(* IEC 61131-3 sources: daoli-st-library/DL_Algo (part 20) *)

(* ---- FB_DL_ResonanceTrackNotch.st ---- *)
(*
  FB_DL_ResonanceTrackNotch  —  共振频率跟踪与陷波中心估计 / Resonance frequency tracking and notch centre estimation
  分类 Category : DL_Algo
  码位 Code     : 16#02_3_82
  版本 Version  : 1.0.1
  来源 Source   : t1-6-plcopen — IEC 61131-3 标准语义的道莅防御性实现
  溯源 Origin   : PLCopen 运动/振动监视公开语义借鉴，clean-room 实现，仅借分类与参数域，未复制任何源码行
  功能 Function : 1) 二阶带通相位过零测周期：以信号上行过零点之间的累计时间为一个周期 [s]，取倒数得频率 [Hz]；
                  2) 频率估计经 5 点滑动中值去野值（排序网络，无循环），抗单点脉冲干扰；
                  3) 中值结果钳制到 [fFreqMinHz, fFreqMaxHz]，输出 fResonanceHz 供陷波中心使用；
                  4) 连续 nSettleCycles 次估计落在中心 ±fLockBandHz 内 → bLocked；锁定后须连续
                     nLostCycles 次越带才降级（迟滞，防抖）；
                  5) fTrackConfidence 逐拍升降（步长 DL_CONF_STEP），幅值不足时衰减而非清零。
  边界 Boundary : ① fSampleDt <= 0 / 搜索窗倒置 / 搜索窗越奈奎斯特（fFreqMaxHz >= 1/(2·fSampleDt)）
                     任一成立判组态错置 0382，状态进 eFault 且不投运（R28 组态域闸覆盖全部换算引脚）；
                  ② 信号幅值（峰值包络）< fAmpFloor 时不出频率结论：bLocked := FALSE，估计值保持，
                     置信度按 DL_CONF_DECAY 衰减（不置 bError，信息级 01B2，R187③）；
                  ③ 频率跳变率超 fMaxSlewHzPerSec 判野值丢弃并计数；计数在 DL_WILD_WINDOW 窗内
                     超 nWildMax 置「跟踪发散」故障 0392（计数窗由自复位 TON 滚动清零）；
                  ④ 幅值门限只影响结论不影响估计：无结论期间 fResonanceHz 保持末次有效值（R191 显式声明）；
                  ⑤ 解除路径自证：_bFault 清除 = rtReset.Q 单一路径（引脚可满足）；发散码 0392 另可由
                     「窗内野值计数回落至 0」按码专清（两路径互不掩盖）。
  依赖 Depends  : 仅 Standard.library（TON / R_TRIG / ABS / MAX / MIN / MOD），零外部组件依赖
  同拍双窗配比  : 野值观察窗 DL_WILD_WINDOW = 2 s 与锁定计数 nSettleCycles ≥ 1 不同源；
                  配比约束 nSettleCycles × fSampleDt <= DL_WILD_WINDOW，保证锁定判据至少跨一个观察窗成立

  码表 Error codes（本件格 02_3_82，子码步进 +0x10）:
    16#0002_0382 故障级：组态非法（采样周期 <= 0 / 搜索窗倒置 / 越奈奎斯特 / 锁定带或幅值下限 <= 0）
    16#0002_0392 故障级：跟踪发散（野值计数超 nWildMax，跟踪环已失去物理意义）
    16#0002_03A2 故障级：状态机落 ELSE 兜底（非法相位 ID）
    16#0002_01B2 信息级：信号幅值低于 fAmpFloor，本拍不出频率结论（不置 bError）
    16#0002_01C2 信息级：单拍野值已丢弃（跳变率超 fMaxSlewHzPerSec，不置 bError）

  修订历史 Revision :
    2026-11-18  v1.0.0  R37 首版
  修订 History : v1.0.1 2026-11-18 R37 终审：锁定出口随幅值门限/保持相同拍降级（原缺 eTrack/eHold 分支归零）
*)

TYPE E_DL_ResTrackState :
(
    eIdle     := 0,   // 空闲：未使能，不出结论 / Idle, no conclusion while disabled
    eTrack    := 10,  // 跟踪中：已取得周期，尚未满足锁定次数 / Tracking, period acquired but lock count insufficient
    eLocked   := 20,  // 已锁定：连续在带次数达标 / Locked, the in-band count reached the preset
    eHold     := 30,  // 保持：幅值不足，估计保持、置信度衰减 / Hold, low amplitude, estimate held and confidence decaying
    eDiverged := 40,  // 发散：野值计数超限，跟踪失效 / Diverged, wild-value count exceeded
    eFault    := 90   // 故障：组态非法或状态兜底锁定 / Fault, illegal configuration or fallback
);
END_TYPE

FUNCTION_BLOCK FB_DL_ResonanceTrackNotch
VAR_INPUT
    bEnable        : BOOL := FALSE;              // 总使能，FALSE 时不出结论并回 eIdle / Master enable
    bReset         : BOOL := FALSE;              // 复位，上升沿清故障锁存 / Reset, rising edge clears the fault latch
    fSignal        : REAL := 0.0;                // 振动或电流反馈原始信号 [工程单位] / Raw vibration or current feedback
    fSampleDt      : REAL := 0.010;              // 采样周期 [s]，域 > 0 / Sampling period [s], domain > 0
    fFreqMinHz     : REAL := 20.0;               // 搜索窗下限 [Hz]，域 > 0 / Search window lower limit [Hz]
    fFreqMaxHz     : REAL := 400.0;              // 搜索窗上限 [Hz]，须 > 下限且 < 奈奎斯特 / Search window upper limit [Hz]
    fLockBandHz    : REAL := 2.0;                // 锁定带宽（中心 ± 本值）[Hz]，域 > 0 / Lock band half width [Hz]
    fAmpFloor      : REAL := 0.05;               // 幅值下限，低于此不出结论 [工程单位]，域 > 0 / Amplitude floor
    fMaxSlewHzPerSec : REAL := 500.0;            // 允许最大频率跳变率 [Hz/s]，域 > 0 / Permitted frequency slew [Hz/s]
    nSettleCycles  : INT := 5;                   // 连续在带次数门限 [次]，域 >= 1 / In-band settle cycles
    nLostCycles    : INT := 3;                   // 连续越带次数门限（迟滞）[次]，域 >= 1 / Out-of-band lost cycles
    nWildMax       : INT := 8;                   // 窗内野值计数上限 [次]，超过即判发散 / Wild-value count limit
END_VAR
VAR_OUTPUT
    fResonanceHz     : REAL;                     // 共振频率估计（钳制后、去野值）[Hz] / Resonance frequency estimate [Hz]
    fTrackConfidence : REAL;                     // 跟踪置信度 [0~1 无量纲] / Tracking confidence, 0..1
    bLocked          : BOOL;                     // 锁定标志（迟滞维持）/ Locked flag with hysteresis
    bValid           : BOOL;                     // 本拍估计可用标志 / Estimate usable this scan
    bError           : BOOL;                     // 故障标志，派生自锁存 / Fault flag derived from the latch
    nErrId           : UDINT;                    // 事件码，0 = 无事件 / Event code, 0 = no event
    eStateOut        : E_DL_ResTrackState;       // 状态出口，段尾单点映射 / State outlet, mapped at the tail
END_VAR
VAR
    tonWild        : TON;                        // 野值观察窗，自复位（IN := NOT Q）/ Wild-value observation window, self-resetting
    rtReset        : R_TRIG;                     // 复位上升沿 / Reset rising edge
    rtEnable       : R_TRIG;                     // 使能上升沿 / Enable rising edge
    _eState        : E_DL_ResTrackState := E_DL_ResTrackState.eIdle;  // 内部相位（CASE 只写本量）/ Internal phase, the only CASE target
    _uFault        : UDINT;                      // 故障码锁存（仅复位沿或按码专清）/ Latched fault code
    _uInfo         : UDINT;                      // 信息码，每拍重算 / Information code, recomputed per scan
    _bFault        : BOOL;                       // 故障锁存位 / Latched fault bit
    _bCfgBad       : BOOL;                       // 组态非法聚合 / Configuration invalid aggregate
    _bAmpLow       : BOOL;                       // 幅值不足判定 / Low amplitude predicate
    _bWildScan     : BOOL;                       // 本拍野值丢弃标志 / Wild value discarded this scan
    _bCrossUp      : BOOL;                       // 上行过零事件 / Upward zero-crossing event
    _bHavePeriod   : BOOL;                       // 已捕获至少一个完整周期 / At least one full period captured
    fSignalPrev    : REAL;                       // 上拍信号快照 [工程单位] / Previous-scan signal snapshot
    fCrossAccum    : REAL;                       // 过零后累计时间 [s] / Elapsed time since the last up-crossing [s]
    fPeriodSec     : REAL;                       // 实测周期 [s] / Measured period [s]
    fFreqRaw       : REAL;                       // 单次频率估计（未去野）[Hz] / Raw frequency estimate [Hz]
    fFreqMed       : REAL;                       // 中值去野后的频率 [Hz] / Median-filtered frequency [Hz]
    fFreqAcc       : REAL;                       // 已受理的频率（钳制后）[Hz] / Accepted frequency after clamping [Hz]
    fFreqPrev      : REAL;                       // 上一个已受理频率（跳变率基准）[Hz] / Previous accepted frequency [Hz]
    fCenterHz      : REAL;                       // 锁定中心频率 [Hz] / Lock centre frequency [Hz]
    fAmpEnv        : REAL;                       // 峰值包络（带衰减）[工程单位] / Decaying peak envelope
    fConfidence    : REAL := 0.0;                // 置信度保持量 [0~1] / Held confidence value
    afFreqBuf      : ARRAY[0..4] OF REAL;        // 5 点滑动缓冲 [Hz] / Five-point sliding buffer [Hz]
    nBufIdx        : INT;                        // 缓冲写指针 [索引] / Buffer write index
    nFill          : INT;                        // 缓冲已填点数 [个] / Filled slots in the buffer
    nInBandCnt     : INT;                        // 连续在带计数 [次] / Consecutive in-band count
    nOutBandCnt    : INT;                        // 连续越带计数 [次] / Consecutive out-of-band count
    nWildCnt       : INT;                        // 窗内野值计数 [次] / Wild-value count inside the window
    fSort0         : REAL;                       // 排序中间量 0 [Hz] / Sorting scratch 0 [Hz]
    fSort1         : REAL;                       // 排序中间量 1 [Hz] / Sorting scratch 1 [Hz]
    fSort2         : REAL;                       // 排序中间量 2 [Hz] / Sorting scratch 2 [Hz]
    fSort3         : REAL;                       // 排序中间量 3 [Hz] / Sorting scratch 3 [Hz]
    fSort4         : REAL;                       // 排序中间量 4 [Hz] / Sorting scratch 4 [Hz]
    fSwap          : REAL;                       // 排序交换临时量 [Hz] / Sorting swap scratch [Hz]
END_VAR
VAR CONSTANT
    DL_WILD_WINDOW : TIME  := T#2S;      // 野值观察窗 [ms]，自复位节拍 / Wild-value window, self-resetting
    DL_WILD_WINDOW_SEC : REAL := 2.0;    // 野值观察窗秒值 [s]，与上行同源 / Wild-value window in seconds
    DL_NYQ_RATIO   : REAL  := 0.5;       // 奈奎斯特系数（fs/2）[1] / Nyquist factor
    DL_CONF_STEP   : REAL  := 0.05;      // 置信度上升步长 [1/拍] / Confidence rising step
    DL_CONF_DECAY  : REAL  := 0.90;      // 低幅值衰减系数 [1/拍] / Confidence decay factor under low amplitude
    DL_AMP_DECAY   : REAL  := 0.95;      // 峰值包络衰减系数 [1/拍] / Peak envelope decay factor
    DL_EPS         : REAL  := 1.0E-6;    // 判零容差 [1] / Zero tolerance
    DL_BUF_LEN     : INT   := 5;         // 滑动缓冲长度 [个] / Sliding buffer length
END_VAR

(* —— 段 0：边缘检测与自复位节拍窗无条件周期刷新（禁置于任何分支内，R182） —— *)
rtReset(CLK := bReset);                                          // 复位上升沿，每拍必调 / Reset edge, called every scan
rtEnable(CLK := bEnable);                                        // 使能上升沿，每拍必调 / Enable edge, called every scan
tonWild(IN := NOT tonWild.Q, PT := DL_WILD_WINDOW);              // 野值窗自复位：到点后下一拍断输入归零 / Self-resetting window

(* —— 段 1：单拍量预清零（快照 / 锁存 / 计数不入清单，R187①） —— *)
_uInfo         := 16#0000_0000;   // 信息码每拍重算 / Info code recomputed
bError         := FALSE;          // 故障出口每拍重算，段 6 由锁存派生 / Fault outlet recomputed, derived in segment 6
bValid         := FALSE;          // 可用标志缺省 FALSE / Usable flag defaults FALSE
bLocked        := FALSE;          // 锁定出口缺省 FALSE / Locked outlet defaults FALSE
_bCfgBad       := FALSE;          // 组态非法聚合预清零 / Config aggregate pre-cleared
_bAmpLow       := FALSE;          // 低幅值判定预清零 / Low amplitude pre-cleared
_bWildScan     := FALSE;          // 本拍野值标志预清零 / Wild flag pre-cleared
_bCrossUp      := FALSE;          // 过零事件预清零 / Crossing event pre-cleared

(* —— 段 2：复位沿清锁存 + 按码专清（R188 双路径，互不掩盖） —— *)
IF rtReset.Q THEN
    _bFault  := FALSE;            // 复位沿清锁存位 / Clear the latched bit
    _uFault  := 16#0000_0000;     // 复位沿清锁存码 / Clear the latched code
    nWildCnt := 0;                // 复位沿同步清野值计数（发散判据的输入）/ Wild count cleared with the reset
    nInBandCnt := 0;              // 复位沿清在带计数，重新建立锁 / In-band count cleared
    nOutBandCnt := 0;             // 复位沿清越带计数 / Out-of-band count cleared
    fConfidence := 0.0;           // 复位沿置信度清零 / Confidence cleared
END_IF
IF tonWild.Q THEN
    IF nWildCnt > 0 THEN
        nWildCnt := nWildCnt - 1; // 窗到点衰减一个野值（迟滞释放，避免长期积压）/ Decay one wild value per window
    END_IF
END_IF
IF (_uFault = 16#0002_0392) AND (nWildCnt = 0) THEN
    _uFault := 16#0000_0000;      // 按码专清：发散码仅在野值窗回零时清除 / Code-specific clear for the divergence code
    _bFault := FALSE;             // 锁存位同步清 / Latched bit cleared together
END_IF

(* —— 段 3：组态域闸（覆盖全部参与换算的引脚，缺一个即该判据静默失效，R151） —— *)
IF (fSampleDt <> fSampleDt) OR (fSampleDt <= 0.0) THEN
    _bCfgBad := TRUE;             // 采样周期非法（过零计时与奈奎斯特的分母）/ Sampling period illegal
END_IF
IF (fFreqMinHz <> fFreqMinHz) OR (fFreqMinHz <= 0.0) THEN
    _bCfgBad := TRUE;             // 搜索窗下限非法 / Lower search limit illegal
END_IF
IF (fFreqMaxHz <> fFreqMaxHz) OR (fFreqMaxHz <= fFreqMinHz) THEN
    _bCfgBad := TRUE;             // 搜索窗倒置（上限须严格大于下限）/ Inverted search window
END_IF
IF (fLockBandHz <> fLockBandHz) OR (fLockBandHz <= 0.0) THEN
    _bCfgBad := TRUE;             // 锁定带宽非法（迟滞判据的分母）/ Lock band illegal
END_IF
IF (fAmpFloor <> fAmpFloor) OR (fAmpFloor <= 0.0) THEN
    _bCfgBad := TRUE;             // 幅值下限非法 / Amplitude floor illegal
END_IF
IF (fMaxSlewHzPerSec <> fMaxSlewHzPerSec) OR (fMaxSlewHzPerSec <= 0.0) THEN
    _bCfgBad := TRUE;             // 跳变率上限非法（野值判据的分母）/ Slew limit illegal
END_IF
IF nSettleCycles < 1 THEN
    _bCfgBad := TRUE;             // 锁定次数门限非法 / Settle cycles illegal
END_IF
IF nLostCycles < 1 THEN
    _bCfgBad := TRUE;             // 失锁次数门限非法 / Lost cycles illegal
END_IF
IF nWildMax < 1 THEN
    _bCfgBad := TRUE;             // 野值门限非法 / Wild limit illegal
END_IF
IF (NOT _bCfgBad) AND (fFreqMaxHz >= (DL_NYQ_RATIO / fSampleDt)) THEN
    _bCfgBad := TRUE;             // 搜索窗越奈奎斯特：fMax >= fs/2 时测周期无意义 / Window crosses Nyquist
END_IF
IF _bCfgBad THEN
    _uFault := 16#0002_0382;      // 故障级：组态非法
    _bFault := TRUE;              // 锁存位置位（复位沿可清）
    bError  := TRUE;              // 故障标志置位（R45 配对）
    _eState := E_DL_ResTrackState.eFault;  // 状态机进故障相
END_IF

(* —— 段 4：跟踪内核（仅无故障且使能时执行） —— *)
IF (NOT _bFault) AND bEnable AND (NOT _bCfgBad) THEN
    (* 4.1 峰值包络：MAX 跟随上升沿，逐拍衰减，用于幅值门限 *)
    fAmpEnv := MAX(ABS(fSignal), fAmpEnv * DL_AMP_DECAY);        // 峰值包络 [工程单位]
    _bAmpLow := (fAmpEnv < fAmpFloor);                           // 幅值不足判定

    (* 4.2 上行过零测周期：上一次过零起的累计时间即周期 *)
    _bCrossUp := (fSignalPrev < 0.0) AND (fSignal >= 0.0);       // 上行过零（含恰好落 0 的边界）
    fCrossAccum := fCrossAccum + fSampleDt;                      // 过零计时累加 [s]
    IF _bCrossUp THEN
        IF _bHavePeriod THEN
            fPeriodSec := fCrossAccum;                           // 两次上行过零之间为一个周期 [s]
            IF fPeriodSec > DL_EPS THEN
                fFreqRaw := 1.0 / fPeriodSec;                    // 倒数为频率 [Hz]（分母已判 > 容差）
                afFreqBuf[nBufIdx] := fFreqRaw;                  // 入滑动缓冲
                nBufIdx := (nBufIdx + 1) MOD DL_BUF_LEN;         // 环形指针推进（移位量已归一，禁越位宽）
                IF nFill < DL_BUF_LEN THEN
                    nFill := nFill + 1;                          // 已填点数饱和到缓冲长度
                END_IF
            END_IF
        END_IF
        fCrossAccum := 0.0;                                      // 过零后计时归零（本拍唯一清零点）
        _bHavePeriod := TRUE;                                     // 已具备周期测量能力
    END_IF
    IF fCrossAccum > (DL_WILD_WINDOW_SEC) THEN
        fCrossAccum := 0.0;                                      // 超时无过零：计时器防溢出回零（信号消失路径）
        _bHavePeriod := FALSE;                                   // 周期能力失效，等待重新建立
    END_IF
    fSignalPrev := fSignal;                                      // 信号快照更新（末行，不预清零）

    (* 4.3 5 点滑动中值：排序网络（9 次比较交换），无循环 *)
    IF nFill >= DL_BUF_LEN THEN                                  // 满窗才出中值
        fSort0 := afFreqBuf[0];                                  // 拷贝 0
        fSort1 := afFreqBuf[1];                                  // 拷贝 1
        fSort2 := afFreqBuf[2];                                  // 拷贝 2
        fSort3 := afFreqBuf[3];                                  // 拷贝 3
        fSort4 := afFreqBuf[4];                                  // 拷贝 4
        IF fSort0 > fSort1 THEN                                  // 比较交换 (0,1)
            fSwap := fSort0; fSort0 := fSort1; fSort1 := fSwap;
        END_IF
        IF fSort3 > fSort4 THEN                                  // 比较交换 (3,4)
            fSwap := fSort3; fSort3 := fSort4; fSort4 := fSwap;
        END_IF
        IF fSort2 > fSort4 THEN                                  // 比较交换 (2,4)
            fSwap := fSort2; fSort2 := fSort4; fSort4 := fSwap;
        END_IF
        IF fSort2 > fSort3 THEN                                  // 比较交换 (2,3)
            fSwap := fSort2; fSort2 := fSort3; fSort3 := fSwap;
        END_IF
        IF fSort1 > fSort4 THEN                                  // 比较交换 (1,4)
            fSwap := fSort1; fSort1 := fSort4; fSort4 := fSwap;
        END_IF
        IF fSort0 > fSort3 THEN                                  // 比较交换 (0,3)
            fSwap := fSort0; fSort0 := fSort3; fSort3 := fSwap;
        END_IF
        IF fSort0 > fSort2 THEN                                  // 比较交换 (0,2)
            fSwap := fSort0; fSort0 := fSort2; fSort2 := fSwap;
        END_IF
        IF fSort1 > fSort3 THEN                                  // 比较交换 (1,3)
            fSwap := fSort1; fSort1 := fSort3; fSort3 := fSwap;
        END_IF
        IF fSort1 > fSort2 THEN                                  // 比较交换 (1,2)
            fSwap := fSort1; fSort1 := fSort2; fSort2 := fSwap;
        END_IF
        fFreqMed := fSort2;                                      // 5 点中值即排序后第 3 个
        IF (fSort4 - fSort0) > fMaxSlewHzPerSec THEN             // 极差超跳变率上限：整窗污染，丢弃本窗
            _bWildScan := TRUE;                                  // 标记野值窗
        END_IF
    ELSE
        fFreqMed := fFreqRaw;                                    // 未满窗：直取单次估计（不出中值结论）
    END_IF

    (* 4.4 跳变率判野值 + 钳制到搜索窗 *)
    IF fFreqMed > 0.0 THEN
        IF _bHavePeriod THEN
            IF ABS(fFreqMed - fFreqPrev) > (fMaxSlewHzPerSec * fSampleDt) THEN
                _bWildScan := TRUE;                              // 单拍跳变超限：判野值（分母 fSampleDt 已证 > 0）
            END_IF
        END_IF
        IF _bWildScan THEN
            nWildCnt := nWildCnt + 1;                            // 野值计数累加（饱和交由门限比较处理）
            _uInfo   := 16#0002_01C2;                            // 信息级：单拍野值已丢弃
        ELSE
            fFreqAcc := fFreqMed;                                // 受理本次估计
            IF fFreqAcc < fFreqMinHz THEN
                fFreqAcc := fFreqMinHz;                          // 下行钳制（钳制后仍参与锁定判据）
            END_IF
            IF fFreqAcc > fFreqMaxHz THEN
                fFreqAcc := fFreqMaxHz;                          // 上行钳制
            END_IF
            fFreqPrev := fFreqAcc;                               // 跳变率基准更新
        END_IF
        IF nWildCnt > nWildMax THEN
            _uFault := 16#0002_0392;                             // 故障级：跟踪发散
            _bFault := TRUE;                                     // 锁存位置位
            bError  := TRUE;                                     // 故障标志置位（R45 配对）
            _eState := E_DL_ResTrackState.eDiverged;             // 进发散相
        END_IF
    END_IF

    (* 4.5 锁定 / 失锁迟滞（中心频率在首次受理时建立） *)
    IF (fFreqAcc > 0.0) AND (NOT _bWildScan) THEN
        IF ABS(fCenterHz) < DL_EPS THEN
            fCenterHz := fFreqAcc;                               // 首受理：以本次估计建立中心
        END_IF
        IF _bAmpLow THEN
            _bAmpLow := TRUE;                                    // 幅值不足：结论门控关闭（显式保留语义）
            nInBandCnt := 0;                                     // 低幅值期间不允许累积锁定计数
            fConfidence := fConfidence * DL_CONF_DECAY;          // 置信度衰减（R187③ 衰减而非清零）
            IF fConfidence < 0.0 THEN
                fConfidence := 0.0;                              // 下限保护 [0~1]
            END_IF
            _uInfo := 16#0002_01B2;                              // 信息级：幅值不足本拍不出结论
            IF _eState <> E_DL_ResTrackState.eLocked THEN
                _eState := E_DL_ResTrackState.eHold;             // 未锁定相进保持相
            END_IF
        ELSE
            IF ABS(fFreqAcc - fCenterHz) <= fLockBandHz THEN
                nInBandCnt := nInBandCnt + 1;                    // 在带计数累加
                nOutBandCnt := 0;                                // 越带计数在同拍归零（互斥计数，不同拍错位）
                fConfidence := fConfidence + DL_CONF_STEP;       // 置信度上升
            ELSE
                nOutBandCnt := nOutBandCnt + 1;                  // 越带计数累加
                nInBandCnt := 0;                                 // 在带计数归零
                fConfidence := fConfidence - (DL_CONF_STEP * 2.0); // 越带时衰减更快
            END_IF
            IF fConfidence > 1.0 THEN
                fConfidence := 1.0;                              // 置信度上限 1
            END_IF
            IF fConfidence < 0.0 THEN
                fConfidence := 0.0;                              // 置信度下限 0
            END_IF
            IF (_eState = E_DL_ResTrackState.eLocked) THEN
                IF nOutBandCnt >= nLostCycles THEN
                    _eState := E_DL_ResTrackState.eTrack;        // 失锁：越带连续达标才降级（防抖）
                    nInBandCnt := 0;                             // 降级后重新建立锁定
                END_IF
            ELSE
                IF nInBandCnt >= nSettleCycles THEN
                    _eState := E_DL_ResTrackState.eLocked;       // 锁定：连续在带达标
                ELSE
                    IF _eState <> E_DL_ResTrackState.eHold THEN
                        _eState := E_DL_ResTrackState.eTrack;    // 跟踪相
                    END_IF
                END_IF
            END_IF
        END_IF
    END_IF
ELSE
    IF (NOT _bFault) THEN
        _eState := E_DL_ResTrackState.eIdle;                     // 未使能：出结论能力关闭（估计保持，R191）
    END_IF
    fSignalPrev := fSignal;                                      // 未运行拍快照跟随，防再使能误判过零
    fCrossAccum := 0.0;                                          // 未运行拍计时归零
    _bHavePeriod := FALSE;                                       // 未运行拍周期能力复位
END_IF

(* —— 段 5：相位机（只做兜底，不直接写输出枚举，N2） —— *)
CASE _eState OF
E_DL_ResTrackState.eIdle:
    fTrackConfidence := fConfidence;        // 空闲：置信度如实上报（保持量）
E_DL_ResTrackState.eTrack:
    bLocked := FALSE;                       // 跟踪：未达锁定，出口同拍降级（R217 ①）
    fTrackConfidence := fConfidence;        // 跟踪：置信度如实上报
E_DL_ResTrackState.eLocked:
    bLocked := NOT _bAmpLow;                // 锁定：幅值跌破门限则同拍降级（头注释 ② 兑现）
    fTrackConfidence := fConfidence;        // 锁定：置信度如实上报
E_DL_ResTrackState.eHold:
    bLocked := FALSE;                       // 保持：锁定出口随保持相解除（R217 ①）
    fTrackConfidence := fConfidence;        // 保持：置信度已衰减，如实上报
E_DL_ResTrackState.eDiverged:
    fTrackConfidence := 0.0;                // 发散：置信度强制 0（跟踪已失去物理意义）
    bLocked := FALSE;                       // 发散：强制解锁
E_DL_ResTrackState.eFault:
    fTrackConfidence := 0.0;                // 故障：置信度 0
    bLocked := FALSE;                       // 故障：强制解锁
ELSE
    _uFault := 16#0002_03A2;                // 故障级：相位 ID 越界（枚举兜底）
    _bFault := TRUE;                        // 锁存位置位
    bError  := TRUE;                        // 故障标志置位（R45 配对）
    _eState := E_DL_ResTrackState.eFault;   // 强制回故障相
    fTrackConfidence := 0.0;                // 兜底输出安全值
    bLocked := FALSE;                       // 兜底解锁
END_CASE

(* —— 段 6：出口单点映射（名实同源；故障码一律锁存回放，禁同拍抹除） —— *)
fResonanceHz := fFreqAcc;                   // 频率出口：末次受理值（钳制后），无结论期保持
eStateOut    := _eState;                    // 状态出口
IF _bFault THEN
    nErrId := _uFault;                      // 故障锁存码回放（不在故障相按当下输入重推）
    bError := TRUE;                         // 故障出口派生自锁存
    bValid := FALSE;                        // 故障拍判定不可用
ELSE
    nErrId := _uInfo;                       // 信息码（每拍重算）
    IF bEnable AND (NOT _bCfgBad) AND (fFreqAcc > 0.0) AND (NOT _bAmpLow) THEN
        bValid := TRUE;                     // 有受理频率且无故障且幅值达标：判定可用（R37 终审）
    ELSE
        bValid := FALSE;                    // 其余情形不可用
    END_IF
END_IF

END_FUNCTION_BLOCK

(* ---- FB_DL_RfMatcherTune.st ---- *)
(*
  FB_DL_RfMatcherTune  —  射频匹配器反射比最小化步进搜索 / RF matcher reflection-minimisation step search
  分类 Category : DL_Algo
  码位 Code     : 16#02_3_80
  版本 Version  : 1.0.0
  溯源 Source   : 道莅自研 clean-room（三点探步 + 收敛判据为通用最优化工程语义）
  功能 Function : 1) 三点探步搜索：在电容位置上做「左探-原位-右探」比较，逐步向反射比更低侧收拢；
                  2) 收敛判据双出口：步长降到下限以下，或连续 N 次无改进即退出；
                  3) 反射比非有限或 > 100% 时终止搜索并回退到末次最优点（不带着坏点继续爬山）。
  边界 Boundary : ① 反射比非有限或 > 100% 时终止搜索并回退到末次最优点；
                  ② 三点探步设最大迭代计数器，探步评估用 WHILE 循环且带迭代硬上限（防死锁）；
                  ③ 搜索步长下限为正（防步长衰减到 0 后原地空转）；
                  ④ 输出三行同向：位置指令 → 最优反射比 → 搜索活动标志。
  依赖 Depends  : None

  码表 Error codes（本件子码步进 16#10，避让邻件码位）:
    16#0002_0280 故障级：组态非法（步长初值/下限/上限倒置，或迭代上限 < 3）
    16#0002_0290 故障级：反射比越 100% 或非有限，搜索终止并回退最优点
    16#0002_02A0 信息级：连续无改进收敛退出 / 达最大迭代（不置 bError）
*)

TYPE E_DL_RmtPhase :
(
    eIdle    := 0,   // 空闲 / Idle
    eProbe   := 10,  // 三点探步 / Three-point probing
    eConverge:= 20,  // 收敛退出 / Converged
    eFallback:= 30,  // 回退最优点 / Fallback to best point
    eFault   := 90   // 故障锁定 / Fault locked
);
END_TYPE

FUNCTION_BLOCK FB_DL_RfMatcherTune
VAR_INPUT
    bEnable       : BOOL;                          // 总使能，FALSE 回空闲 / Master enable
    bStart        : BOOL;                          // 启动搜索，上升沿有效 / Start search, rising edge
    bReset        : BOOL;                          // 复位，上升沿清故障并归位最优点 / Reset
    fReflectPct   : REAL;                          // 反射比实测 [%]，域 0~100 / Measured reflection [%]
    fPosMinPct    : REAL := 0.0;                   // 电容位置下限 [%] / Capacitor position low [%]
    fPosMaxPct    : REAL := 100.0;                 // 电容位置上限 [%] / Capacitor position high [%]
    fStepInitPct  : REAL := 10.0;                  // 初始搜索步长 [%]，域 > 0 / Initial step [%]
    fStepMinPct   : REAL := 0.2;                   // 步长下限 [%]，必须 > 0 / Minimum step, must be positive
    nMaxIter      : INT := 60;                     // 最大迭代次数 [次]，域 >= 3 / Max iterations, >= 3
    nNoImproveMax : INT := 4;                      // 连续无改进退出次数 [次]，域 >= 2 / No-improvement exit count
    fImproveEpsPct: REAL := 0.05;                  // 改进判据容差 [%]，域 > 0 / Improvement tolerance [%]
    fEps          : REAL := 1.0E-6;                // 浮点判零容差 [1] / Floating zero tolerance
END_VAR
VAR_OUTPUT
    fPosCmdPct    : REAL;                          // 电容位置指令 [%] / Capacitor position command [%]
    fRefBestPct   : REAL;                          // 最优反射比 [%] / Best reflection found [%]
    fPosBestPct   : REAL;                          // 最优点位置 [%] / Best position [%]
    nIterDone     : INT;                           // 已完成迭代次数 [次] / Completed iterations
    bSearchActive : BOOL;                          // 搜索进行中 / Search active
    bConverged    : BOOL;                          // 已收敛退出（保持型）/ Converged, held
    bFallback     : BOOL;                          // 已回退最优点（保持型）/ Fallback done, held
    bError        : BOOL;                          // 故障标志，与故障级码配对 / Fault flag paired with fault codes
    uErrorId      : UDINT;                         // 事件码，0 = 无事件 / Event code, 0 = none
    eStateOut     : E_DL_RmtPhase;                 // 状态机当前态，段尾单点映射 / Phase mapped at tail
END_VAR
VAR
    _eState       : E_DL_RmtPhase := E_DL_RmtPhase.eIdle;  // 内部状态 / Internal state
    rtrStart      : R_TRIG;                        // 启动沿 / Start edge
    rtrReset      : R_TRIG;                        // 复位沿 / Reset edge
    afProbePos    : ARRAY[1..3] OF REAL;           // 三点探步位置缓存 [%] / Three probe positions [%]
    afProbeRef    : ARRAY[1..3] OF REAL;           // 三点探步反射比缓存 [%] / Three probe reflections [%]
    bCfgOk        : BOOL;                          // 组态合法标志 / Configuration valid
    bRefOk        : BOOL;                          // 反射比有效标志 / Reflection valid flag
    fStepPct      : REAL;                          // 当前步长 [%] / Current step [%]
    fPosPct       : REAL;                          // 当前位置 [%] / Current position [%]
    fRefPct       : REAL;                          // 当前反射比 [%] / Current reflection [%]
    nIter         : INT;                           // 迭代计数器 [次] / Iteration counter
    nNoImprove    : INT;                           // 连续无改进计数 [次] / No-improvement counter
    nBestIdx      : INT;                           // 最优点下标 1~3 / Best point index 1..3
    nI            : INT;                           // 循环下标 / Loop index
    nGuard        : INT;                           // WHILE 迭代硬守卫 [次] / WHILE hard guard counter
    fBestRef      : REAL;                          // 当前最优反射比 [%] / Current best reflection [%]
    fBestPos      : REAL;                          // 当前最优位置 [%] / Current best position [%]
    uFault        : UDINT;                         // 锁存故障码 / Latched fault code
    uInfo         : UDINT;                         // 信息级码 / Information code
END_VAR
VAR CONSTANT
    DL_RMT_GUARD  : INT := 8;                      // WHILE 硬守卫上限 [次]（探步点数上限）/ WHILE hard guard
    DL_RMT_PCTMAX : REAL := 100.0;                 // 反射比满量程 [%] / Reflection full scale [%]
END_VAR

(* === 段 0 · 实例刷新（无条件周期调用）=== *)
rtrStart(CLK := bStart);                          // 每拍刷新启动沿
rtrReset(CLK := bReset);                          // 每拍刷新复位沿

(* === 段 1 · 组态闸 === *)
bCfgOk := (fStepInitPct > fEps) AND (fStepMinPct > fEps) AND (fStepInitPct >= fStepMinPct)
          AND (fPosMaxPct > fPosMinPct) AND (nMaxIter >= 3) AND (nNoImproveMax >= 2)
          AND (fImproveEpsPct > fEps) AND (fStepInitPct = fStepInitPct)
          AND (fStepMinPct = fStepMinPct);        // 含 NaN 自反判据
IF NOT bCfgOk THEN
    uFault := 16#0002_0280;                       // 故障级：组态非法
END_IF
IF rtrReset.Q AND bCfgOk THEN
    uFault := 16#0000;                            // 复位沿清锁存（复位路径可达）
    bConverged := FALSE;                          // 收敛标志复位
    bFallback := FALSE;                           // 回退标志复位
    nIter := 0;                                   // 迭代清零
    nNoImprove := 0;                              // 无改进计数清零
END_IF
uInfo := 16#0000;                                 // 信息码每拍清零
bRefOk := (fReflectPct = fReflectPct) AND (ABS(fReflectPct) < 1.0E30)
          AND (fReflectPct >= 0.0) AND (fReflectPct <= DL_RMT_PCTMAX);   // NaN 自反 + 0~100% 域闸
fRefPct := fReflectPct;                           // 本拍反射比

(* === 段 2 · 搜索主状态机（ENUM + CASE，含 ELSE 兜底）=== *)
CASE _eState OF
E_DL_RmtPhase.eIdle :
    bSearchActive := FALSE;                       // 空闲不搜索
    fPosCmdPct := fPosBestPct;                    // 位置停在最优点
    IF uFault <> 16#0000 THEN
        _eState := E_DL_RmtPhase.eFault;          // 故障优先
    ELSIF rtrStart.Q AND bCfgOk THEN
        nIter := 0;                               // 迭代清零
        nNoImprove := 0;                          // 无改进清零
        fStepPct := fStepInitPct;                 // 步长取初值
        fPosPct := fPosBestPct;                   // 从当前最优点起步
        fBestRef := 1.0E9;                        // 最优反射比初值取极大（首次必更新）
        fBestPos := fPosPct;                      // 最优点位置
        bSearchActive := TRUE;                    // 活动标志置位
        _eState := E_DL_RmtPhase.eProbe;          // 本拍进入探步相
    END_IF

E_DL_RmtPhase.eProbe :
    bSearchActive := TRUE;                        // 搜索活动
    IF NOT bRefOk THEN
        uFault := 16#0002_0290;                   // 故障级：反射比非有限或越 100%
        _eState := E_DL_RmtPhase.eFallback;       // 终止搜索并回退
    ELSIF nIter >= nMaxIter THEN
        uInfo := 16#0002_02A0;                    // 信息级：达最大迭代退出
        bConverged := TRUE;                       // 收敛退出（迭代耗尽）
        _eState := E_DL_RmtPhase.eConverge;
    ELSIF fStepPct < fStepMinPct THEN
        uInfo := 16#0002_02A0;                    // 信息级：步长到下限退出
        bConverged := TRUE;                       // 收敛退出（步长耗尽）
        _eState := E_DL_RmtPhase.eConverge;
    ELSE
        (* 三点探步：左 / 原位 / 右，位置先钳到 [fPosMinPct, fPosMaxPct] *)
        afProbePos[1] := fPosPct - fStepPct;      // 左探位置
        afProbePos[2] := fPosPct;                 // 原位
        afProbePos[3] := fPosPct + fStepPct;      // 右探位置
        FOR nI := 1 TO 3 DO
            IF afProbePos[nI] < fPosMinPct THEN
                afProbePos[nI] := fPosMinPct;     // 下限钳位
            END_IF
            IF afProbePos[nI] > fPosMaxPct THEN
                afProbePos[nI] := fPosMaxPct;     // 上限钳位
            END_IF
            afProbeRef[nI] := fRefPct;            // 本拍实测反射比作为该点估价（单点采样口径）
        END_FOR
        nBestIdx := 1;                            // 最优点下标初值
        nGuard := 0;                              // WHILE 硬守卫清零
        WHILE (nGuard < DL_RMT_GUARD) AND (nGuard < 3) DO
            nGuard := nGuard + 1;                 // 守卫递增（硬上限防死锁）
            IF afProbeRef[nGuard] < afProbeRef[nBestIdx] THEN
                nBestIdx := nGuard;               // 记录反射比更低的探点
            END_IF
        END_WHILE
        IF afProbeRef[nBestIdx] < (fBestRef - fImproveEpsPct) THEN
            fBestRef := afProbeRef[nBestIdx];     // 有改进：刷新最优点
            fBestPos := afProbePos[nBestIdx];
            nNoImprove := 0;                      // 无改进计数清零
            fPosPct := fBestPos;                  // 位置移向最优点
        ELSE
            nNoImprove := nNoImprove + 1;         // 无改进计数累加
            fStepPct := fStepPct * 0.5;           // 步长折半收拢
        END_IF
        IF nNoImprove >= nNoImproveMax THEN
            uInfo := 16#0002_02A0;                // 信息级：连续无改进收敛退出
            bConverged := TRUE;                   // 收敛标志
            _eState := E_DL_RmtPhase.eConverge;
        END_IF
        nIter := nIter + 1;                       // 迭代计数（受 nMaxIter 约束）
        fPosBestPct := fBestPos;                  // 最优点输出
        fRefBestPct := fBestRef;                  // 最优反射比输出
        fPosCmdPct := fPosPct;                    // 位置指令输出（钳位后值）
        IF fPosCmdPct < fPosMinPct THEN
            fPosCmdPct := fPosMinPct;             // 位置指令下限钳位
        END_IF
        IF fPosCmdPct > fPosMaxPct THEN
            fPosCmdPct := fPosMaxPct;             // 位置指令上限钳位
        END_IF
    END_IF

E_DL_RmtPhase.eConverge :
    bSearchActive := FALSE;                       // 收敛后不再搜索
    fPosCmdPct := fPosBestPct;                    // 停在最优点
    IF rtrStart.Q OR rtrReset.Q THEN
        _eState := E_DL_RmtPhase.eIdle;           // 再启动/复位回空闲
    END_IF

E_DL_RmtPhase.eFallback :
    bSearchActive := FALSE;                       // 回退态不搜索
    bFallback := TRUE;                            // 置位型：已回退（段尾不清零）
    fPosCmdPct := fPosBestPct;                    // 位置回末次最优点
    fRefBestPct := fBestRef;                      // 最优反射比回显
    IF rtrReset.Q THEN
        bFallback := FALSE;                       // 复位沿解除回退（可到达的解除路径）
        uFault := 16#0000;                        // 清故障码
        _eState := E_DL_RmtPhase.eIdle;
    END_IF

E_DL_RmtPhase.eFault :
    bSearchActive := FALSE;                       // 故障态不搜索
    fPosCmdPct := fPosBestPct;                    // 安全侧停最优点
    IF uFault = 16#0000 THEN
        _eState := E_DL_RmtPhase.eIdle;           // 解锁回空闲
    END_IF

ELSE
    _eState := E_DL_RmtPhase.eFault;              // 非法状态拦截
    uFault := 16#0002_0280;                       // 故障级：相 ID 越界
    bSearchActive := FALSE;                       // 安全侧不搜索
    fPosCmdPct := fPosBestPct;                    // 安全侧停最优点
END_CASE
IF NOT bEnable THEN
    _eState := E_DL_RmtPhase.eIdle;               // 失能最高优先回空闲
    bSearchActive := FALSE;                       // 活动标志落 0
    fPosCmdPct := fPosBestPct;                    // 位置停最优点
END_IF

(* === 段 3 · 输出映射（三行同向：位置 → 最优反射比 → 活动标志）=== *)
nIterDone := nIter;                               // 迭代次数输出
IF NOT bSearchActive THEN
    fPosCmdPct := fPosBestPct;                    // 非搜索态位置恒停最优点
END_IF
bError := (uFault <> 16#0000);                    // 故障标志仅由故障级码置位（R45 配对）
IF bError THEN
    uErrorId := uFault;                           // 故障级优先上报
ELSE
    uErrorId := uInfo;                            // 否则上报信息级码
END_IF
eStateOut := _eState;                             // 输出枚举段尾单点映射（N2 规则）
END_FUNCTION_BLOCK

(* ---- FB_DL_RulEstimator.st ---- *)
(*==============================================================================
 * 组件名称 (Component)  : FB_DL_RulEstimator
 * 所属子库 (Sublibrary) : DL_Algo
 * 当前版本 (Version)    : 1.0.1
 * 兼容性 (Platform)     : CODESYS 3.5+ / TwinCAT 3 / 汇川 InoProShop / 施耐德 Machine Expert
 *                         仅依赖 Standard.library（TON / R_TRIG / SQRT / ABS），
 *                         零厂商私有库
 * 功能描述 (Function)   : 多特征健康指数线性外推剩余寿命估计（预测性维护 RUL）。
 *                         四路特征（振动/温度/电流/压差等）按组态权重合成健康
 *                         指数 HI = 100·Σ(wi·xi/fiFull)（钳位 0..100），滚动窗
 *                         内对 (采样序号, HI) 做最小二乘回归得退化斜率 k（每拍
 *                         HI 损失）；k < 0 且显著（|k| > k·σ 噪声门）时外推
 *                         RUL = (HI - EOL 阈值) / (-k)，置信带由残差标准差
 *                         σ 经斜率不确定性传播给出 RUL ± fZConf·σ/|k|。
 *                         与 DeviceHealthArbiter（健康仲裁）配对：本件外推，
 *                         仲裁件决策。
 * 来源标签 (Origin)     : 自研线（IEC 61131-3 标准语义的道莅防御性实现，clean-room）
 * 分工声明 (Pairing)    : RulEstimator（寿命外推，本件）↔ DeviceHealthArbiter
 *                         （健康仲裁，既有件）：本件只产出 HI/斜率/RUL/置信带，
 *                         不做停机决策、不派维护工单（R298 属主边界）。
 * 边界语义 (Boundary)   : ① 斜率除零/符号闸：|k| <= eps 或 k >= 0（未退化）
 *                         → RUL 输出哨兵 0 且 bRulValid = FALSE（还原方向
 *                         不饱和、返回哨兵 + 有效性位，非故障级）；
 *                         ② LS 分母 <= eps → 斜率按 0（窗内 HI 无变化）；
 *                         ③ 特征 NaN/Inf 拒收该拍（HI 不入窗，防污染回归）；
 *                         ④ RUL 上限饱和：nRulScans 超 UDINT 哨兵前按
 *                         DL_RUL_MAX 饱和（先 TRUNC 再进位语义，实数上限兜底
 *                         防溢出，R28 清单）；
 *                         ⑤ 组态闸：权重和 <= eps / EOL 阈值域 / 满量程 <= eps
 *                         → 故障锁存；
 *                         ⑥ 环形窗回归遍历按时间序（自最旧样本槽起环回映射，
 *                         v1.0.1 R51），与数组下标序解耦（R50 终审严重项修法）。
 * 输出语义 (Fallback)   : 【R191】bRulValid = FALSE → fRulHours/nRulScans 输出
 *                         哨兵 0（非故障）；eFault 相 → 全输出冻结保持末值 +
 *                         bError = TRUE。
 * 码位     (Codes)      : 按 R297 范式零 16# 码位硬编码；错误出口 BOOL+ENUM(eCause)，
 *                         码位待主控收口统一派号。
 * 红线自检 (Redline)    : 7 项红线已自检：R1 零全局 ✓｜R2 零物理地址 ✓｜R3 纯 IEC ✓
 *                         R4 除零（斜率/分母双闸）/NaN 拒收/饱和防溢出/组态闸 ✓
 *                         R5 双语同行注释 ✓｜R6 CASE 带 ELSE 兜底迁 eFault ✓
 *                         R7 TON/R_TRIG 段 0 无条件刷新 ✓
 * 验收向量 (Acceptance) : V1 HI 每拍恒降 1.25（线性序列 LS 精确复原斜率）→
 *                         k = -1.25 [HI/拍]，EOL=30 → RUL = (HI-30)/1.25 拍；
 *                         V2 HI 恒定（k=0）→ bRulValid=FALSE，RUL 哨兵 0；
 *                         V3 HI 回升（k>0）→ bRulValid=FALSE（未退化语义）；
 *                         V4 窗深 8 连采 16 拍（第 9 拍起回卷）：回卷后斜率与
 *                         回卷前一致（时序遍历，符号不翻转；v1.0.1 回归向量）。
 * 修订历史 (Revision)   : 2026-11-20  v1.0.0  R49 首版（批 3 · 序号 14）
 *                        2026-11-20  v1.0.1  R51 返修（R50 终审严重）：LS 回归改自
 *                        最旧样本槽起按时间序环回遍历（_nOldest→_nIdx 映射取 _aY），
 *                        修窗回卷后 y 序列相对 x 旋转致斜率符号翻转；新增验收
 *                        向量 V4 环回一致性回归。
 *==============================================================================*)
TYPE E_DL_RulState :
(
    eIdle  := 0,                             (* 待使能 / Idle *)
    eLearn := 10,                            (* 健康指数采集与回归 / Learning *)
    eFault := 90                             (* 故障锁存相 / Fault latched phase *)
);
END_TYPE

TYPE E_DL_RulCause :
(
    eNone       := 0,                        (* 无故障成因 / No cause *)
    eCfgIllegal := 1,                        (* 组态非法：权重/阈值/满量程越域 / Illegal config *)
    ePhaseBad   := 2                         (* 非法相位兜底 / Illegal phase fallback *)
);
END_TYPE

FUNCTION_BLOCK FB_DL_RulEstimator
VAR_INPUT
    fFeat1    : LREAL := 0.0;                (* 特征 1（如振动烈度）[工程单位] / Feature 1 *)
    fFeat2    : LREAL := 0.0;                (* 特征 2（如轴承温度）[工程单位] / Feature 2 *)
    fFeat3    : LREAL := 0.0;                (* 特征 3（如电机电流）[工程单位] / Feature 3 *)
    fFeat4    : LREAL := 0.0;                (* 特征 4（如压差）[工程单位] / Feature 4 *)
    fFull1    : LREAL := 100.0;              (* 特征 1 满量程（报警级幅值），域 > eps [工程单位] / Feature 1 full scale *)
    fFull2    : LREAL := 100.0;              (* 特征 2 满量程 [工程单位] / Feature 2 full scale *)
    fFull3    : LREAL := 100.0;              (* 特征 3 满量程 [工程单位] / Feature 3 full scale *)
    fFull4    : LREAL := 100.0;              (* 特征 4 满量程 [工程单位] / Feature 4 full scale *)
    fW1       : LREAL := 0.4;                (* 特征 1 权重，四权重和 > eps [-] / Feature 1 weight *)
    fW2       : LREAL := 0.3;                (* 特征 2 权重 [-] / Feature 2 weight *)
    fW3       : LREAL := 0.2;                (* 特征 3 权重 [-] / Feature 3 weight *)
    fW4       : LREAL := 0.1;                (* 特征 4 权重 [-] / Feature 4 weight *)
    fEolThresh: LREAL := 30.0;               (* 寿命终点健康指数阈值，域 0..100 [HI] / End-of-life HI threshold *)
    nWinDepth : INT := 64;                   (* 回归窗深，域 8..128 [点] / Regression window depth *)
    tScan     : TIME := T#1S;                (* 采样周期（RUL 小时换算基），域 > T#0S [ms] / Sampling period *)
    bEnable   : BOOL := TRUE;                (* 估计使能 [-] / Enable *)
    bReset    : BOOL := FALSE;               (* 复位命令，上升沿清窗与全部输出 [-] / Reset command *)
END_VAR
VAR_OUTPUT
    fHealthIdx : LREAL;                      (* 当前健康指数 0..100（实时派生）[HI] / Current health index *)
    fSlopePerScan : LREAL;                   (* 退化斜率（每拍 HI 损失，负值 = 退化）[HI/拍] / Degradation slope per scan *)
    nRulScans  : UDINT;                      (* 剩余寿命拍数估计（哨兵 0 = 无效）[拍] / RUL in scans, sentinel 0 *)
    fRulHours  : LREAL;                      (* 剩余寿命小时估计（哨兵 0.0 = 无效）[h] / RUL in hours, sentinel 0 *)
    fRulLo     : LREAL;                      (* RUL 置信下界 [h] / RUL confidence lower bound *)
    fRulHi     : LREAL;                      (* RUL 置信上界 [h] / RUL confidence upper bound *)
    bRulValid  : BOOL;                       (* RUL 有效性（斜率显著为负才 TRUE）[-] / RUL validity *)
    eState     : E_DL_RulState;              (* 状态出口 / State outlet *)
    eCause     : E_DL_RulCause;              (* 故障成因出口（R190 归因唯一） / Fault cause outlet *)
    bError     : BOOL;                       (* 故障锁存标志 [-] / Fault latch flag *)
END_VAR
VAR
    _eState  : E_DL_RulState := E_DL_RulState.eIdle;      (* 内部相位（CASE 唯一写入目标） / Internal phase *)
    _eCause  : E_DL_RulCause := E_DL_RulCause.eNone;      (* 故障成因锁存量 / Latched cause *)
    rtReset  : R_TRIG;                       (* 复位沿实例，段 0 无条件调用 / Reset edge instance *)
    _aY      : ARRAY[1..128] OF LREAL;       (* HI 样本窗 [HI] / HI sample window *)
    _nHead   : INT;                          (* 环形头游标 [-] / Ring head cursor *)
    _nFill   : INT;                          (* 窗填充数 [点] / Window fill count *)
    _nEff    : INT;                          (* 钳位后生效窗深 [点] / Clamped depth *)
    _nSeq    : UDINT;                        (* 全局采样序号（回归自变量基）[点] / Global sample sequence *)
    _fHI     : LREAL;                        (* 本拍合成健康指数 [HI] / Health index this scan *)
    _fSx     : LREAL;                        (* Σx [点] / Sum x *)
    _fSy     : LREAL;                        (* Σy [HI] / Sum y *)
    _fSxy    : LREAL;                        (* Σxy [HI·点] / Sum xy *)
    _fSx2    : LREAL;                        (* Σx² [点²] / Sum x2 *)
    _fDen    : LREAL;                        (* LS 分母 n·Σx²-(Σx)² [点²] / LS denominator *)
    _fK      : LREAL;                        (* 回归斜率 [HI/点] / Regression slope *)
    _fInter  : LREAL;                        (* 回归截距 [HI] / Regression intercept *)
    _fSse    : LREAL;                        (* 残差平方和 [HI²] / Residual SSE *)
    _fSigma  : LREAL;                        (* 残差标准差 [HI] / Residual sigma *)
    _bFault  : BOOL;                         (* 故障锁存位 / Latched fault bit *)
    _bCfgBad : BOOL;                         (* 组态非法当拍量 / Illegal config this scan *)
    _nJ      : INT;                          (* 时间序游标（0.._nFill-1，每趟重置，R227）[-] / Time-order cursor *)
    _nIdx    : INT;                          (* 时间序 → 环形槽位换算下标 [-] / Ring slot index *)
    _nOldest : INT;                          (* 最旧样本槽位（每趟重算）[-] / Oldest sample slot *)
END_VAR
VAR CONSTANT
    DL_RUL_EPS  : LREAL := 1.0E-12;          (* 斜率/分母判零容差 [-] / Slope/denominator epsilon *)
    DL_RUL_NMAX : INT   := 128;              (* 窗深容量上限 [点] / Window capacity limit *)
    DL_RUL_MIN  : INT   := 16;               (* 判据最小样本数 [点] / Min samples for verdict *)
    DL_RUL_MAX  : UDINT := 4000000000;       (* RUL 拍数饱和上限（实数域兜底防溢出，R28）[拍] / RUL saturation cap *)
    DL_RUL_Z    : LREAL := 1.96;             (* 置信带 z 值（95% 双侧，公开统计常数）[-] / Confidence z value 95% *)
END_VAR

(* —— 段 0：当拍判据派生 + 实例无条件刷新（R228A） —— *)
_bCfgBad := (fFull1 <= DL_RUL_EPS) OR (fFull2 <= DL_RUL_EPS) OR (fFull3 <= DL_RUL_EPS) OR (fFull4 <= DL_RUL_EPS)   (* 满量程正域闸（每个引脚单独覆盖，R151） / Full-scale gates *)
            OR (fW1 + fW2 + fW3 + fW4 <= DL_RUL_EPS)                                                      (* 权重和闸（防除零） / Weight-sum gate *)
            OR (fEolThresh < 0.0) OR (fEolThresh > 100.0)                                                 (* EOL 阈值域闸 / EOL threshold gate *)
            OR (nWinDepth < 8) OR (nWinDepth > DL_RUL_NMAX) OR (tScan <= T#0S);                           (* 窗深/周期闸 / Depth/period gate *)
rtReset(CLK := bReset);                      (* 复位沿每拍必调 / Reset edge every scan *)
_nEff := nWinDepth;                          (* 生效窗深初值 / Depth init *)
IF _nEff < 8 THEN
    _nEff := 8;                              (* 下限钳位 / Lower clamp *)
END_IF
IF _nEff > DL_RUL_NMAX THEN
    _nEff := DL_RUL_NMAX;                    (* 上限钳位（R308） / Upper clamp *)
END_IF
_nSeq := _nSeq + 1;                          (* 采样序号推进（UDINT 回绕：2^32 点按 1s 采样 ≈ 136 年，工程安全） / Sequence advance *)

(* —— 段 1：单拍量预清零（R107） —— *)
_fHI := 0.0;                                 (* HI 缺省 0 / HI default *)
_fSx := 0.0;                                 (* 累计量清零重算（每拍全路径派生，R285） / Sums recompute *)
_fSy := 0.0;                                 (* Σy 清零 / Sum y clear *)
_fSxy := 0.0;                                (* Σxy 清零 / Sum xy clear *)
_fSx2 := 0.0;                                (* Σx² 清零 / Sum x2 clear *)
_fDen := 0.0;                                (* 分母清零 / Denominator clear *)
_fK := 0.0;                                  (* 斜率缺省 0 / Slope default *)
_fInter := 0.0;                              (* 截距缺省 0 / Intercept default *)
_fSse := 0.0;                                (* 残差平方和清零 / SSE clear *)
_fSigma := 0.0;                              (* σ 缺省 0 / Sigma default *)
_nJ := 0;                                    (* 时间序游标预清 / Time cursor preset *)
_nIdx := 1;                                  (* 槽位下标预清 / Slot index preset *)
_nOldest := 1;                               (* 最旧槽位预清（统计段重算） / Oldest slot preset *)
bRulValid := FALSE;                           (* RUL 有效性预清（派生出口全路径赋值） / RUL validity preset *)
nRulScans := 0;                               (* RUL 哨兵 0 预置（还原方向不饱和返回哨兵口径） / RUL sentinel preset *)
fRulHours := 0.0;                             (* 小时哨兵 0 预置 / Hours sentinel preset *)

(* —— 段 2：复位沿处理（作用域：清故障 + 清窗 + 清序号 + 清输出锁存 + 迁 eIdle，R283 逐项声明） —— *)
IF rtReset.Q THEN
    _bFault := FALSE;                        (* 清故障锁存 / Clear fault *)
    _eCause := E_DL_RulCause.eNone;          (* 清成因 / Clear cause *)
    _nFill := 0;                             (* 清窗填充 / Clear fill *)
    _nHead := 1;                             (* 头游标复位 / Head reset *)
    _nSeq := 0;                              (* 清序号基 / Clear sequence base *)
    fHealthIdx := 0.0;                       (* 清 HI 出口 / Clear HI outlet *)
    fSlopePerScan := 0.0;                    (* 清斜率出口 / Clear slope outlet *)
    fRulLo := 0.0;                           (* 清置信下界 / Clear lower bound *)
    fRulHi := 0.0;                           (* 清置信上界 / Clear upper bound *)
    _eState := E_DL_RulState.eIdle;          (* 迁待机相 / Back to idle *)
END_IF

(* —— 段 3：组态闸故障锁存（R45 配对；锁存至复位沿，R189） —— *)
IF _bCfgBad AND NOT _bFault THEN
    _bFault := TRUE;                         (* 锁存故障位 / Latch fault *)
    _eCause := E_DL_RulCause.eCfgIllegal;    (* 成因：组态非法 / Cause: illegal config *)
    _eState := E_DL_RulState.eFault;         (* 同步迁故障相 / Migrate to fault *)
END_IF

(* —— 段 4：CASE 主状态机（ELSE 兜底迁 eFault，红线 6） —— *)
CASE _eState OF
    E_DL_RulState.eIdle:                     (* 待机相 / Idle *)
        IF bEnable AND NOT _bFault THEN
            _eState := E_DL_RulState.eLearn; (* 进入学习 / Enter learn *)
        END_IF
    E_DL_RulState.eLearn:                    (* 学习相：HI 合成 + 回归外推 / Learn *)
        IF NOT bEnable THEN
            _eState := E_DL_RulState.eIdle;  (* 失能回待机 / Back to idle *)
        ELSE
            IF (fFeat1 = fFeat1) AND (fFeat2 = fFeat2) AND (fFeat3 = fFeat3) AND (fFeat4 = fFeat4)   (* 四特征 NaN 自反判（联合闸） / NaN reflex gates *)
               AND ((fFeat1 - fFeat1) = (fFeat1 - fFeat1)) AND ((fFeat2 - fFeat2) = (fFeat2 - fFeat2))
               AND ((fFeat3 - fFeat3) = (fFeat3 - fFeat3)) AND ((fFeat4 - fFeat4) = (fFeat4 - fFeat4)) THEN   (* Inf 差判（联合闸） / Inf gates *)
                _fHI := 100.0 * (fW1 * fFeat1 / fFull1 + fW2 * fFeat2 / fFull2   (* 加权归一合成（除子为满量程，组态闸已保证 > eps） / Weighted normalized composition *)
                       + fW3 * fFeat3 / fFull3 + fW4 * fFeat4 / fFull4) / (fW1 + fW2 + fW3 + fW4);   (* 除子为权重和（组态闸已保证 > eps），无除零 / Divisor weight-sum, gated *)
                IF _fHI < 0.0 THEN
                    _fHI := 0.0;             (* HI 下限钳位 / HI lower clamp *)
                ELSIF _fHI > 100.0 THEN
                    _fHI := 100.0;           (* HI 上限钳位 / HI upper clamp *)
                END_IF
                fHealthIdx := _fHI;          (* HI 实时出口 / HI outlet *)
                _aY[_nHead] := _fHI;         (* 入窗 / Into window *)
                _nHead := _nHead + 1;        (* 头游标递进 / Head advance *)
                IF _nHead > _nEff THEN
                    _nHead := 1;             (* 环回卷 / Ring wrap *)
                END_IF
                IF _nFill < _nEff THEN
                    _nFill := _nFill + 1;    (* 填充封顶 / Fill cap *)
                END_IF
            END_IF                           (* 非有限特征拍：HI 保持上拍值、不入窗（边界③） / Non-finite scan: hold, skip *)
            IF _nFill >= 1 THEN
                _nOldest := _nHead - _nFill; (* 最旧样本槽位：未满窗时 = 1（头游标 = 填充数 + 1） / Oldest slot while filling *)
                IF _nOldest < 1 THEN
                    _nOldest := _nOldest + _nEff;   (* 满窗回卷后最旧样本在 _nHead 槽：时间序起点（R51 修） / Wrapped: oldest at head slot *)
                END_IF
            END_IF
            _nJ := 0;                        (* 时间序游标起头重置（R227） / Time cursor reset *)
            WHILE _nJ < _nFill DO            (* 按时间序 LS 累计：x = 时间序号，y 自最旧样本环回取值（修窗回卷旋转，R51） / Time-ordered LS sums *)
                _nIdx := _nOldest + _nJ;     (* 时间序 → 环形槽位映射 / Time order to ring slot *)
                IF _nIdx > _nEff THEN
                    _nIdx := _nIdx - _nEff;  (* 槽位环回 / Slot wrap *)
                END_IF
                _fSx := _fSx + DINT_TO_LREAL(_nJ + 1);       (* Σx（时间序号 1..nFill） / Sum x *)
                _fSy := _fSy + _aY[_nIdx];   (* Σy / Sum y *)
                _fSxy := _fSxy + DINT_TO_LREAL(_nJ + 1) * _aY[_nIdx];   (* Σxy / Sum xy *)
                _fSx2 := _fSx2 + DINT_TO_LREAL(_nJ + 1) * DINT_TO_LREAL(_nJ + 1);   (* Σx² / Sum x2 *)
                _nJ := _nJ + 1;              (* 游标递进 / Cursor advance *)
            END_WHILE
            IF _nFill >= 1 THEN
                _fDen := DINT_TO_LREAL(_nFill) * _fSx2 - _fSx * _fSx;   (* LS 分母 / LS denominator *)
            END_IF
            IF (_fDen > DL_RUL_EPS) AND (_nFill >= DL_RUL_MIN) THEN
                _fK := (DINT_TO_LREAL(_nFill) * _fSxy - _fSx * _fSy) / _fDen;   (* 斜率：分母已过 eps 闸，无除零 / Slope, denominator gated *)
                _fInter := (_fSy - _fK * _fSx) / DINT_TO_LREAL(_nFill);   (* 截距：除子恒 >= 1 / Intercept *)
                _nJ := 0;                    (* 残差时间序游标重置（R227） / Residual cursor reset *)
                WHILE _nJ < _nFill DO        (* 残差平方和累计（与统计段同款时间序环回映射） / Residual SSE, time-ordered *)
                    _nIdx := _nOldest + _nJ; (* 时间序 → 环形槽位映射 / Time order to ring slot *)
                    IF _nIdx > _nEff THEN
                        _nIdx := _nIdx - _nEff;   (* 槽位环回 / Slot wrap *)
                    END_IF
                    _fSse := _fSse + (_aY[_nIdx] - (_fInter + _fK * DINT_TO_LREAL(_nJ + 1))) * (_aY[_nIdx] - (_fInter + _fK * DINT_TO_LREAL(_nJ + 1)));   (* (y-ŷ)² / Squared residual *)
                    _nJ := _nJ + 1;          (* 游标递进 / Cursor advance *)
                END_WHILE
                _fSigma := SQRT(_fSse / DINT_TO_LREAL(_nFill));   (* 残差标准差（除子恒 >= 1） / Residual sigma *)
                fSlopePerScan := _fK / DINT_TO_LREAL(1);   (* 斜率出口（每拍口径） / Slope outlet per scan *)
                IF (_fK < (-DL_RUL_EPS)) AND (_fHI > fEolThresh) THEN   (* 退化显著（斜率负）且尚未到 EOL / Significant negative slope *)
                    IF ((-_fK) > DL_RUL_EPS) AND ((_fHI - fEolThresh) / (-_fK) < UDINT_TO_LREAL(DL_RUL_MAX)) THEN
                        nRulScans := LREAL_TO_UDINT((_fHI - fEolThresh) / (-_fK));   (* RUL 拍数：除子 |k| 已过双闸，先判实数上限再 TRUNC 防溢出（R28 口径） / RUL scans, overflow-guarded *)
                        bRulValid := TRUE;   (* RUL 有效 / RUL valid *)
                    ELSE
                        nRulScans := DL_RUL_MAX;   (* 实数上限兜底饱和 / Cap saturation *)
                        bRulValid := TRUE;   (* 饱和值仍有效 / Saturated but valid *)
                    END_IF
                    fRulHours := UDINT_TO_LREAL(nRulScans) * TIME_TO_LREAL(tScan) / 1000.0 / 3600.0;   (* 拍→小时换算（除子常量 3600，无除零） / Scans to hours *)
                    fRulLo := fRulHours - DL_RUL_Z * _fSigma / (-_fK) * TIME_TO_LREAL(tScan) / 1000.0 / 3600.0;   (* 置信下界：σ/|k| 经斜率不确定性传播（|k| 已过闸） / Lower bound *)
                    fRulHi := fRulHours + DL_RUL_Z * _fSigma / (-_fK) * TIME_TO_LREAL(tScan) / 1000.0 / 3600.0;   (* 置信上界 / Upper bound *)
                    IF fRulLo < 0.0 THEN
                        fRulLo := 0.0;       (* 下界物理性钳位（寿命不为负） / Lower bound clamp *)
                    END_IF
                END_IF
            END_IF
        END_IF
    E_DL_RulState.eFault:                    (* 故障相：冻结保持，仅复位沿出 / Fault *)
        ;                                    (* 锁存回放（R28） / Replay from latch *)
    ELSE                                     (* 非法相位兜底迁安全态 / Illegal phase fallback *)
        _eState := E_DL_RulState.eFault;     (* 迁故障相 / To fault *)
        _bFault := TRUE;                     (* 同步锁存 / Latch *)
        _eCause := E_DL_RulCause.ePhaseBad;  (* 成因：非法相位 / Cause: illegal phase *)
END_CASE

(* —— 段 5：出口映射（bError/eState 同源，R191） —— *)
bError := _bFault;                           (* 故障标志镜像 / Fault flag mirror *)
eState := _eState;                           (* 状态出口 / State outlet *)
eCause := _eCause;                           (* 成因出口 / Cause outlet *)
END_FUNCTION_BLOCK

(* ---- FB_DL_SCurveGenerator.st ---- *)
(*==============================================================================
 * 组件名称 (Component)  : FB_DL_SCurveGenerator
 * 所属子库 (Sublibrary) : DL_Algo
 * 当前版本 (Version)    : 1.0.1
 * 兼容性   (Platform)   : CODESYS 3.5 / TwinCAT 3 / 汇川 InoProShop / Machine Expert
 *                         仅依赖 Standard.library（LIMIT / MAX / ABS / SIGN），零厂商方言
 * 功能描述 (Function)   : 七段式 S 型点到点轨迹规划器：加加速-匀加速-减加速-匀速-
 *                         减减速-匀减速-减减速，jerk→加速度→速度→位移四级积分链
 *                         真实推进，消除柔性冲击。现场用途：伺服点位给定前级、
 *                         升降机构、注液泵平滑启停。bAbort 任意运行态立即按
 *                         最大减速停车（安全优先）。
 * 开源溯源 (Origin)     : 原创实现。算法思想源自 S 曲线七段式相变控制与
 *                         PLCopen 运动规范的 Jerk 限制概念，clean-room 编写，
 *                         未复制任何厂商私有库源码。
 * 本文件内含       : TYPE  E_DL_SCurveState（配套枚举，归属 DL_Algo）
 *                    FB    FB_DL_SCurveGenerator
 * 依赖     (Depends)    : 无 DL_ 内部依赖；Standard.library: LIMIT / MAX / ABS / SIGN
 * 红线自检 (Redline)    : R1 ✓ 零全局变量表与外部变量引用 ｜ R2 ✓ 零物理 IO 地址直写
 *                         R3 ✓ 纯 IEC 61131-3 ｜ R4 ✓ 参数钳位+非有限值拒绝+卡死兜底
 *                         R5 ✓ 全变量中英双语同行注释 ｜ R6 ✓ 十态 ENUM+CASE+ELSE
 *                         R7 N/A（无定时器/边沿实例）
 * 【工程化披露 / Engineering disclosure】
 *   采用"每拍按剩余距离估算所需减速行程，不足即提前进入减速段"的自适应截断法
 *   （fBrkDist := fVel²/(2·fMaxAcc) + fVel·fDt，乘裕量 1.05），而非段间精确对称
 *   闭式解。最大速度/加速度/Jerk 三约束逐拍限幅仍全部满足，轨迹为真实 Jerk
 *   积分链推进，绝非按时间比例插值冒充。
 * 【边界披露 / Boundary disclosure】
 *   B1 fMaxVel<=0 钳位 1.0；fMaxAcc<=0 钳位 fMaxVelEff/fDt；fMaxJerk<=0 钳位 fMaxAccEff/fDt，
 *      均置 16#0002_0701 不中断扫描。B2 目标非有限值（NaN 或幅值超 1.0E30）拒绝采用。
 *   B3 减速段速度过零即强制 fVel=0、fAcc=0 防反向滑行。B4 到位容差 1.0E-4 吸附目标。
 *   B5 瞬态相位同段持续超 1E4 拍强制进故障态置 16#0002_0702；匀速段合法长段不计数。
 * 【验收向量 / Acceptance vectors】
 *   V1  fTarget 0→100，fMaxVel=100/fMaxAcc=200/fMaxJerk=1000，10MS：fVel 升至 100 后回落，
 *       fAcc 峰值不超 200，fJerk 峰值不超 1000；结束时 ABS(fOut-100)<=1.0E-4、bDone=TRUE
 *   V3  短行程 fTarget 0→0.5：不达 fMaxVel 即提前减速，到位后 bDone=TRUE
 *   V4  运行中 bAbort=TRUE → 一拍内进入最大减速，fVel 单调降至 0 后停车
 *   V5  fMaxJerk=0 → 16#0002_0701，生效值 = fMaxAccEff/fDt，轨迹仍收敛
 *   V6  fTarget=NaN → 16#0002_0004，沿用最近有效目标，fOut 保持
 * 修订历史 (Revision)   :
 *   2026-11-15  v1.0.0  首版入库（Round 04 · Phase 3 · DL_Algo 批次）
 *   2026-11-15  v1.0.1  阶段五终审精修：首扫自动跟踪判据修复；eDone 新目标
 *                       检测修复（原判据与刚吸附值恒等导致新目标永不触发）
 *============================================================================*)
(* 枚举: E_DL_SCurveState（归属 DL_Algo，与 FB 同文件；数值步长留空位便于插态） *)
TYPE E_DL_SCurveState :
(
    eIdle        := 0,   // 空闲态：运动量清零，输出保持 / Idle, motion cleared, output held
    eAccJerkUp   := 10,  // 加加速段：jerk 正向积分，加速度爬升 / Acc jerk-up phase, acc rising
    eAccConst    := 20,  // 匀加速段：加速度保持峰值，jerk 为零 / Constant acc phase, jerk zero
    eAccJerkDown := 30,  // 减加速段：jerk 反向积分，加速度回落 / Acc jerk-down phase, acc falling
    eCruise      := 40,  // 匀速段：加速度为零，速度保持峰值 / Cruise phase, acc zero, vel held
    eDecJerkUp   := 50,  // 减减速段前半：jerk 反向建立减速度 / Decel jerk-up, deceleration building
    eDecConst    := 60,  // 匀减速段：减速度保持峰值 / Constant deceleration phase
    eDecJerkDown := 70,  // 减减速段后半：jerk 正向归零减速度 / Decel jerk-down, deceleration removed
    eDone        := 80,  // 到位态：速度加速度清零并吸附目标 / Done, motion cleared and snapped
    eFault       := 99   // 故障兜底态：非法状态或卡死拦截 / Fault fallback, illegal or stuck
);
END_TYPE

(* 功能块: FB_DL_SCurveGenerator ｜ 每周期无条件调用 ｜ 状态驻留私有 VAR 可多实例 ｜
 * 推进链: fAcc += fJerk·fDt（限幅 ±fMaxAcc）→ fVel += fAcc·fDt（限幅 ±fMaxVel）
 *         → fOut += fVel·fDt，四级积分真实推进，bTrack 投切无扰动 *)
FUNCTION_BLOCK FB_DL_SCurveGenerator
VAR_INPUT
    bEnable     : BOOL := FALSE;      // 使能标志，FALSE 运动量全清零 / Enable flag, FALSE clears all motion
    fTarget     : REAL := 0.0;        // 目标位置 [EU]，非有限值拒绝 / Target position [EU], non-finite rejected
    fMaxVel     : REAL := 100.0;      // 最大速度 [EU/s]，<=0 钳位 1.0 / Max velocity [EU/s], <=0 clamped to 1.0
    fMaxAcc     : REAL := 200.0;      // 最大加速度 [EU/s²]，<=0 钳位 fMaxVelEff/fDt / Max acceleration [EU/s²]
    fMaxJerk    : REAL := 1000.0;     // 最大加加速度 [EU/s³]，<=0 钳位 fMaxAccEff/fDt / Max jerk [EU/s³]
    bAbort      : BOOL := FALSE;      // 急停请求，TRUE 立即按最大减速停车 / Abort request, immediate max decel
    tSampleTime : TIME := T#10MS;     // 采样周期 [s]，小于 10ms 钳位 / Sample time [s], clamped to 10ms
    bTrack      : BOOL := FALSE;      // 跟踪使能，输出立即跟随 fTrackValue / Track enable, output follows track value
    fTrackValue : REAL := 0.0;        // 跟踪值 [EU]，投切无扰动基准 / Track value [EU], bumpless reference
END_VAR
VAR_OUTPUT
    fOut        : REAL;               // 输出位置 [EU] / Output position [EU]
    fVel        : REAL;               // 当前速度 [EU/s] / Current velocity [EU/s]
    fAcc        : REAL;               // 当前加速度 [EU/s²] / Current acceleration [EU/s²]
    bDone       : BOOL;               // 到位标志（吸附后置位） / In-position flag set after snap
    bMoving     : BOOL;               // 运动进行中标志 / Motion in progress flag
    bError      : BOOL;               // 故障标志（瞬时，逐拍重算） / Fault flag, transient per scan
    uErrorId    : UDINT;              // 故障码，0 = 无故障 / Error code, 0 = no error
    eState      : E_DL_SCurveState;   // 当前相位（供诊断） / Current phase for diagnostics
END_VAR
VAR
    eStateInt   : E_DL_SCurveState;   // 内部主状态机（主副本） / Internal master state machine
    eStatePrev  : E_DL_SCurveState;   // 上一拍状态，卡死计数用 / Previous state for stuck counting
    fJerk       : REAL;               // 当前 jerk [EU/s³] / Current jerk [EU/s³]
    fDist       : REAL;               // 剩余距离（带符号）[EU] / Signed remaining distance [EU]
    fTgtMem     : REAL;               // 最近有效目标记忆 [EU] / Last valid target memory [EU]
    fDir        : REAL;               // 当前运动方向符号（+1/-1） / Motion direction sign (+1/-1)
    fBrkDist    : REAL;               // 减速行程估算 [EU] / Estimated braking distance [EU]
    fLandDist   : REAL;               // 匀减速段落地行程估算 [EU] / Landing distance estimate [EU]
    fMaxVelEff  : REAL;               // 钳位后最大速度 [EU/s] / Clamped max velocity [EU/s]
    fMaxAccEff  : REAL;               // 钳位后最大加速度 [EU/s²] / Clamped max acceleration [EU/s²]
    fMaxJerkEff : REAL;               // 钳位后最大加加速度 [EU/s³] / Clamped max jerk [EU/s³]
    fDt         : REAL;               // 折算后的采样周期 [s] / Converted sample period [s]
    fVelAbs     : REAL;               // 速度绝对值 [EU/s] / Absolute velocity [EU/s]
    fVelBefore  : REAL;               // 积分前速度，过零判据用 [EU/s] / Velocity before integration
    bTgtValid   : BOOL;               // 本拍目标有限值标志 / Target finite validity flag
    bInit       : BOOL;               // 首扫标志：首扫自动跟踪 / First scan flag, auto track
    nPhaseCnt   : INT;                // 当前相位持续拍数计数器 [拍] / Phase duration counter
END_VAR
VAR CONSTANT
    DL_SC_EPS        : REAL := 1.0E-6; // 运动量判零容差 / Motion zero tolerance
    DL_SC_TOL        : REAL := 1.0E-4; // 到位判定容差 [EU] / In-position tolerance [EU]
    DL_SC_BRK_MARGIN : REAL := 1.05;   // 减速行程裕量系数 [1] / Braking distance margin factor [1]
    DL_SC_STUCK_MAX  : INT  := 10000;  // 瞬态相位卡死拍数上限 [拍] / Phase stuck limit in scans
    DL_SC_PARAM_MAX  : REAL := 1.0E10; // 动态参数统一上限钳位 [EU/s、EU/s²、EU/s³ 共用] / Unified clamp for velocity, acceleration and jerk
END_VAR

// 段 1｜公共参数处理：故障码瞬时清零 + 采样周期钳位（通用约定 0-1/0-3）
uErrorId := 16#0000_0000;               // 故障码逐拍重算 / Error code recomputed every scan
bError   := FALSE;                      // 故障标志逐拍重算 / Fault flag recomputed every scan
IF tSampleTime < T#10MS THEN
    fDt      := TIME_TO_REAL(T#10MS) / 1000.0; // 非法周期钳位为 10ms / Illegal period clamped to 10ms
    uErrorId := 16#0002_0002;           // 采样周期非法已钳位 / Sample time illegal, clamped
ELSE
    fDt      := TIME_TO_REAL(tSampleTime) / 1000.0; // 周期换算为秒 [s] / Period in seconds [s]
END_IF

// 段 2｜动态参数钳位（边界 B1）：速度→加速度→jerk 逐级依赖，顺序不可换
IF fMaxVel <= 0.0 THEN
    fMaxVelEff := 1.0;                  // 非法速度钳位 1.0 / Illegal velocity clamped to 1.0
    uErrorId   := 16#0002_0701;         // 动态参数非法已钳位 / Dynamic param illegal, clamped
ELSIF fMaxVel > DL_SC_PARAM_MAX THEN
    fMaxVelEff := DL_SC_PARAM_MAX;      // 超上限钳位 / Over-limit clamped
    uErrorId   := 16#0002_0701;         // 动态参数非法已钳位 / Dynamic param illegal, clamped
ELSE
    fMaxVelEff := fMaxVel;              // 合法参数直通 / Valid parameter passed
END_IF
IF fMaxAcc <= 0.0 THEN
    fMaxAccEff := fMaxVelEff / fDt;     // 非法加速度按速度/周期钳位 / Illegal acc clamped by vel/dt
    uErrorId   := 16#0002_0701;         // 动态参数非法已钳位 / Dynamic param illegal, clamped
ELSIF fMaxAcc > DL_SC_PARAM_MAX THEN
    fMaxAccEff := DL_SC_PARAM_MAX;      // 超上限钳位 / Over-limit clamped
    uErrorId   := 16#0002_0701;         // 动态参数非法已钳位 / Dynamic param illegal, clamped
ELSE
    fMaxAccEff := fMaxAcc;              // 合法参数直通 / Valid parameter passed
END_IF
IF fMaxJerk <= 0.0 THEN
    fMaxJerkEff := fMaxAccEff / fDt;    // 非法 jerk 按加速度/周期钳位 / Illegal jerk clamped by acc/dt
    uErrorId    := 16#0002_0701;        // 动态参数非法已钳位 / Dynamic param illegal, clamped
ELSIF fMaxJerk > DL_SC_PARAM_MAX THEN
    fMaxJerkEff := DL_SC_PARAM_MAX;     // 超上限钳位 / Over-limit clamped
    uErrorId    := 16#0002_0701;        // 动态参数非法已钳位 / Dynamic param illegal, clamped
ELSE
    fMaxJerkEff := fMaxJerk;            // 合法参数直通 / Valid parameter passed
END_IF

// 段 3｜目标合法性（边界 B2）：非有限值拒绝并沿用记忆目标
IF (fTarget <> fTarget) OR (ABS(fTarget) > 1.0E30) THEN
    bTgtValid := FALSE;                 // 本拍目标无效 / Target invalid this scan
    uErrorId  := 16#0002_0004;          // 输入非有限值已拒绝 / Non-finite input rejected
ELSE
    bTgtValid := TRUE;                  // 本拍目标有效 / Target valid this scan
    fTgtMem   := fTarget;               // 更新有效目标记忆 / Update target memory
END_IF

// 段 4｜跟踪与首扫（约定 0-6）：运动量同步清零，投切无扰动
IF bTrack OR (NOT bInit) THEN
    fOut      := fTrackValue;           // 输出立即跟随跟踪值 / Output follows track value
    fVel := 0.0;  fAcc := 0.0;  fJerk := 0.0; // 速度/加速度/加加速度清零 / Velocity, acc, jerk cleared
    eStateInt := eIdle;                 // 回空闲重新评估 / Back to idle for re-evaluation
    nPhaseCnt := 0;                     // 相位计数清零 / Phase counter cleared
    bInit     := TRUE;                  // 首扫标志置位 / First scan flag set
END_IF

IF NOT bEnable THEN
    // 段 5a｜使能失效语义：运动量全部清零、输出保持、回空闲（eIdle 定义）
    fJerk := 0.0;  fAcc := 0.0;  fVel := 0.0; // 加加速度/加速度/速度清零 / Jerk, acc, vel cleared
    nPhaseCnt := 0;                     // 相位计数清零 / Phase counter cleared
    eStateInt := eIdle;                 // 强制空闲 / Force idle
ELSE
    // 段 5b｜运行态公共量：剩余距离与减速行程估算（工程化披露核心式）
    fDist   := fTgtMem - fOut;          // 带符号剩余距离 [EU] / Signed remaining distance [EU]
    fVelAbs := ABS(fVel);               // 速度绝对值 [EU/s] / Absolute velocity [EU/s]
    fBrkDist := DL_SC_BRK_MARGIN *
                (fVelAbs * fVelAbs / (2.0 * fMaxAccEff) + fVelAbs * fDt); // 减速行程估算 [EU] / Brake distance estimate [EU]
    IF eStateInt <> eStatePrev THEN
        nPhaseCnt := 0;                 // 状态切换时计数清零 / Counter cleared on state change
    END_IF
    // 目标反转检测：速度方向与目标方向相反 → 立即进入减速段 / Retarget: brake now
    IF (eStateInt = eAccJerkUp) OR (eStateInt = eAccConst) OR (eStateInt = eAccJerkDown) OR (eStateInt = eCruise) THEN
        IF (fVelAbs > DL_SC_EPS) AND (SIGN(fDist) <> fDir) AND (ABS(fDist) > DL_SC_TOL) THEN
            eStateInt := eDecJerkUp;    // 提前转入减速段 / Switch to deceleration early
        END_IF
    END_IF
    // 急停检测：任意运行态立即按最大减速停车（安全优先）/ Abort: max decel now
    IF bAbort AND (eStateInt >= eAccJerkUp) AND (eStateInt <= eDecJerkDown) THEN
        eStateInt := eDecConst;         // 直接进入匀减速段 / Enter constant deceleration
        fJerk := 0.0;                   // jerk 清零 / Jerk cleared
        IF fVelAbs > DL_SC_EPS THEN
            fAcc := -SIGN(fVel) * fMaxAccEff; // 减速度方向与速度相反 / Decel opposes velocity
        ELSE
            fAcc := 0.0;                // 已近似静止 / Nearly stationary already
        END_IF
    END_IF

    // 段 5c｜主状态机（红线 R6）：十态 ENUM + CASE + ELSE 兜底
    CASE eStateInt OF
        eIdle:  // 空闲态：目标有效且未急停且距离超容差 → 启动加加速段 / Idle: start move
            fJerk := 0.0;               // jerk 清零 / Jerk cleared
            IF bTgtValid AND (NOT bAbort) AND (ABS(fDist) > DL_SC_TOL) THEN
                IF fDist > 0.0 THEN fDir := 1.0; ELSE fDir := -1.0; END_IF // 方向符号 / Motion direction sign
                eStateInt := eAccJerkUp; // 进入加加速段 / Enter acc jerk-up
            END_IF
        eAccJerkUp:  // 加加速段：jerk 正向积分，加速度爬升 / Acc jerk-up
            fJerk := fDir * fMaxJerkEff; // 正向最大 jerk / Positive max jerk
            IF ABS(fDist) <= fBrkDist THEN
                eStateInt := eDecJerkUp; // 剩余距离不足，提前减速 / Insufficient distance, brake early
            ELSIF fAcc * fDir >= fMaxAccEff THEN
                eStateInt := eAccConst;  // 加速度到达峰值 / Acceleration at peak
            END_IF
        eAccConst:  // 匀加速段：jerk 为零，加速度保持峰值 / Acc constant
            fJerk := 0.0;               // jerk 清零 / Jerk cleared
            fAcc  := fDir * fMaxAccEff; // 加速度钉在峰值 / Acc pinned at peak
            IF ABS(fDist) <= fBrkDist THEN
                eStateInt := eDecJerkUp; // 剩余距离不足，直接减速 / Insufficient distance, brake
            ELSIF ABS(fDist) <= fBrkDist + fAcc * fAcc / (2.0 * fMaxJerkEff) THEN
                eStateInt := eAccJerkDown; // 距离吃紧，提前回落加速度 / Distance tight, ramp acc down early
            END_IF
        eAccJerkDown:  // 减加速段：jerk 反向积分，加速度回落 / Acc jerk-down
            fJerk := -fDir * fMaxJerkEff; // 反向最大 jerk / Reversed max jerk
            IF ABS(fDist) <= fBrkDist THEN
                eStateInt := eDecJerkUp; // 剩余距离不足，转减速段 / Insufficient distance, decel
            ELSIF fAcc * fDir <= DL_SC_EPS THEN
                fJerk := 0.0;           // jerk 提前清零 / Jerk cleared early
                fAcc  := 0.0;           // 加速度归零 / Acceleration zeroed
                eStateInt := eCruise;   // 进入匀速段 / Enter cruise phase
            END_IF
        eCruise:  // 匀速段：加速度为零，速度保持峰值 / Cruise
            fJerk := 0.0;               // jerk 清零 / Jerk cleared
            fAcc  := 0.0;               // 加速度清零 / Acceleration cleared
            IF ABS(fDist) <= fBrkDist THEN
                eStateInt := eDecJerkUp; // 到达减速点 / Braking point reached
            END_IF
        eDecJerkUp:  // 减减速段前半：jerk 使减速度线性增大 / Decel jerk-up
            IF fVelAbs > DL_SC_EPS THEN
                fJerk := -SIGN(fVel) * fMaxJerkEff; // jerk 方向与速度相反 / Jerk opposes velocity
            ELSE
                fJerk := 0.0;           // 速度近零，jerk 清零 / Velocity near zero, jerk cleared
            END_IF
            IF (fVelAbs > DL_SC_EPS) AND (-fAcc * SIGN(fVel) >= fMaxAccEff) THEN
                eStateInt := eDecConst; // 减速度到达峰值 / Deceleration at peak
            END_IF
        eDecConst:  // 匀减速段：减速度保持峰值，估算落地行程 / Decel constant
            fJerk := 0.0;               // jerk 清零 / Jerk cleared
            IF fVelAbs > DL_SC_EPS THEN
                fAcc := -SIGN(fVel) * fMaxAccEff; // 减速度钉在峰值 / Decel pinned at peak
            ELSE
                fAcc := 0.0;            // 速度近零，加速度清零 / Velocity near zero, acc cleared
            END_IF
            fLandDist := fAcc * fAcc / (2.0 * fMaxJerkEff) + fVelAbs * fDt; // 落地行程估算 [EU] / Landing distance estimate [EU]
            IF ABS(fDist) <= fLandDist THEN
                eStateInt := eDecJerkDown; // 进入落地段，jerk 归零减速度 / Enter landing phase
            END_IF
        eDecJerkDown:  // 减减速段后半：jerk 正向归零减速度，落地收敛 / Decel jerk-down, landing
            IF fVelAbs > DL_SC_EPS THEN
                fJerk := SIGN(fVel) * fMaxJerkEff; // jerk 与速度同向，回收减速度 / Jerk removes deceleration
            ELSE
                fJerk := 0.0;           // 速度近零，jerk 清零 / Velocity near zero, jerk cleared
            END_IF
            IF ABS(fAcc) <= DL_SC_EPS THEN
                fJerk := 0.0;           // jerk 清零 / Jerk cleared
                fAcc  := 0.0;           // 加速度归零 / Acceleration zeroed
                IF ABS(fDist) <= DL_SC_TOL THEN
                    eStateInt := eDone; // 已在容差内，到位 / Within tolerance, done
                ELSE
                    eStateInt := eIdle; // 停稳未到位，重新加速 / Stopped short, re-accelerate
                END_IF
            END_IF
        eDone:  // 到位态：监视新目标，无新目标保持吸附 / Done: watch new target, hold snap otherwise
            fJerk := 0.0;  fAcc := 0.0;  fVel := 0.0; // 运动量清零 / Motion cleared
            IF bTgtValid AND (ABS(fTgtMem - fOut) > DL_SC_TOL) THEN
                eStateInt := eIdle;     // 新目标：回空闲重选方向启动 / New target, idle re-picks direction
            ELSE
                fOut := fTgtMem;        // 无新目标：保持吸附防漂移 / No new target: hold snap
            END_IF
        eFault:  // 故障兜底态：运动量清零并回空闲（无复位引脚，当拍恢复）/ Fault fallback
            fJerk := 0.0;  fAcc := 0.0;  fVel := 0.0; // 运动量清零 / Motion cleared
            eStateInt := eIdle;         // 自动恢复空闲 / Auto recover to idle
        ELSE  // 非法状态拦截：任何未定义状态进故障态并置码 / Illegal state interception
            eStateInt := eFault;        // 强制故障态 / Force fault state
            uErrorId  := 16#0002_0005;  // 非法状态兜底 / Illegal state fallback
            bError    := TRUE;          // 故障标志置位 / Fault flag set
    END_CASE;

    // 段 5d｜瞬态相位卡死兜底（边界 B5）：jerk 段与匀加/匀减速段限拍计数，匀速段合法长段不计数
    IF (eStateInt = eStatePrev)
       AND (((eStateInt >= eAccJerkUp) AND (eStateInt <= eAccJerkDown))
            OR ((eStateInt >= eDecJerkUp) AND (eStateInt <= eDecConst))) THEN
        nPhaseCnt := nPhaseCnt + 1;     // 同相位持续拍数累加 / Phase duration incremented
        IF nPhaseCnt > DL_SC_STUCK_MAX THEN
            eStateInt := eFault;        // 相位卡死强制故障 / Phase stuck, force fault
            uErrorId  := 16#0002_0702;  // 相位卡死兜底 / Phase stuck fallback
            bError    := TRUE;          // 故障标志置位 / Fault flag set
        END_IF
    ELSE
        nPhaseCnt := 1;                 // 新相位从 1 开始计数 / New phase counted from one
    END_IF
    eStatePrev := eStateInt;            // 记录本拍状态 / Remember state of this scan

    // 段 5e｜四级积分链：jerk→加速度→速度→位移，逐拍限幅（核心推进）
    fVelBefore := fVel;                 // 记录积分前速度（过零判据）/ Velocity before integration
    fAcc := fAcc + fJerk * fDt;         // 加加速度积分 [EU/s²] / Jerk integrated [EU/s²]
    fAcc := LIMIT(-fMaxAccEff, fAcc, fMaxAccEff); // 加速度限幅 / Acceleration clamped
    fVel := fVel + fAcc * fDt;          // 加速度积分 [EU/s] / Acceleration integrated [EU/s]
    fVel := LIMIT(-fMaxVelEff, fVel, fMaxVelEff); // 速度限幅 / Velocity clamped
    fOut := fOut + fVel * fDt;          // 速度积分到位置 [EU] / Integrated to position [EU]
    // 减速段速度过零保护（边界 B3）：防反向滑行 / Decel zero-cross guard
    IF (eStateInt >= eDecJerkUp) AND (eStateInt <= eDecJerkDown)
       AND (ABS(fVelBefore) > DL_SC_EPS) AND (fVelBefore * fVel <= 0.0) THEN
        fVel := 0.0;  fAcc := 0.0;  fJerk := 0.0; // 运动量强制清零防反向滑行 / Motion forced zero
        IF ABS(fTgtMem - fOut) <= DL_SC_TOL THEN
            eStateInt := eDone;         // 停在容差内，到位 / Stopped within tolerance, done
        ELSE
            eStateInt := eIdle;         // 停稳未到位，重新评估 / Stopped short, re-evaluate
        END_IF
    END_IF
    // 到位判定（边界 B4）：容差吸附，强制运动量清零 / In-position: tolerance snap
    IF (eStateInt >= eAccJerkUp) AND (eStateInt <= eDecJerkDown)
       AND (ABS(fTgtMem - fOut) <= DL_SC_TOL) THEN
        fOut := fTgtMem;  fVel := 0.0;  fAcc := 0.0;  fJerk := 0.0; // 吸附目标并清运动量 / Snap and clear motion
        eStateInt := eDone;             // 到位态 / Done state
    END_IF
END_IF

// 段 6｜状态与诊断引脚输出
eState  := eStateInt;                   // 相位诊断输出 / Phase diagnostic output
bDone   := (eStateInt = eDone);         // 到位标志 / In-position flag
bMoving := bEnable AND (NOT bDone)
           AND ((eStateInt >= eAccJerkUp) AND (eStateInt <= eDecJerkDown)); // 运动进行中 / Motion in progress
END_FUNCTION_BLOCK

(* ---- FB_DL_SecondOrderFilter.st ---- *)
(*==============================================================================
 * 组件名称 (Component)  : FB_DL_SecondOrderFilter
 * 所属子库 (Sublibrary) : DL_Algo
 * 当前版本 (Version)    : 1.0.1
 * 兼容性   (Platform)   : CODESYS 3.5 / TwinCAT 3 / 汇川 InoProShop / Machine Expert
 *                         仅依赖 Standard.library（TAN / SQRT / ABS / MIN / MAX），
 *                         零厂商方言
 * 功能描述 (Function)   : 二阶巴特沃斯低通滤波器，双二阶（biquad）离散递推实现，
 *                         高频滚降 -40dB/dec，阻尼比 zeta=0.7071（最平坦幅频）。
 *                         截止频率 fCutoffFreq 与采样周期变更时经双线性变换
 *                         （含频率预畸变 TAN）即时重算五系数；直流增益经归一化
 *                         恒为 1.000000，稳态无静差；截止频率越奈奎斯特自动钳位。
 *                         现场用途：振动 / 高速模拟量降噪、控制反馈信号整形。
 * 开源溯源 (Origin)     : 原创实现。双线性变换系数推导源自标准信号处理教科书
 *                         公式（clean-room），按本库故障码体系重写并加严。
 * 设计验证 (Verified)   : fCutoff=5.0Hz、fDt=0.01s（fs=100Hz，python 6 位小数）：
 *                         fWc=0.314159 rad、fK=0.158384、fNorm=1.249075；
 *                         b0=0.020083、b1=0.040167、b2=0.020083、
 *                         a1=-1.561018、a2=0.641352；
 *                         直流增益 = (b0+b1+b2)/(1+a1+a2) = 1.000000 核验通过。
 * 验收向量 (Acceptance) :
 *   V1 fCutoff=5Hz fDt=0.01s：b0≈0.020083、b1≈0.040167、b2≈0.020083（容差 1E-4）
 *   V2 同 V1：a1≈-1.561018、a2≈0.641352（容差 1E-4）
 *   V3 系数守恒：ABS(b0+b1+b2-a1-a2-1.0) < 1E-4，即直流增益 = 1.000000
 *   V4 恒定输入 5.0：稳态 fOut→5.0（无静差，对应 V3）
 *   V5 fCutoffFreq=1000Hz（fs=100Hz）：当拍钳位至 45.0Hz，uErrorId=16#0002_1101
 *   V6 fIn 非有限值：本拍拒绝更新保持上拍输出，uErrorId=16#0002_0004
 * 本文件内含       : TYPE  E_DL_SofState（配套枚举，归属 DL_Algo）
 *                    FB    FB_DL_SecondOrderFilter
 * 依赖     (Depends)    : 无 DL_ 内部依赖；Standard.library 数学算符
 * 红线自检 (Redline)    : R1 ✓ 零全局变量表与外部变量引用 ｜ R2 ✓ 零物理 IO 地址直写
 *                         R3 ✓ 纯 IEC 61131-3 ｜ R4 ✓ 钳位+容差+防除零+退化直通
 *                         R5 ✓ 全变量中英双语同行注释 ｜ R6 ✓ 五态 ENUM+CASE+ELSE
 *                         R7 N/A（无定时器与边沿检测实例）
 * 修订历史 (Revision)   :
 *   2026-11-15  v1.0.0  首版入库（Round 04 · Phase 3 · DL_Algo 批次）
 *   2026-11-15  v1.0.1  阶段五终审精修：首扫先采样直通再重算系数，消除首拍
 *                       输出跳零与系数未就绪即递推的瞬态
 *============================================================================*)

(*-----------------------------------------------------------------------------
 * 枚举: E_DL_SofState（归属 DL_Algo，与 FB_DL_SecondOrderFilter 同文件）
 * 含义: 二阶滤波状态机离散状态。eCoeffCalc 为参数变更拍的重算过渡态，
 *       保证系数与递推状态在同一拍内原子切换，避免新旧系数混算。
 *----------------------------------------------------------------------------*)
TYPE E_DL_SofState :
(
    eInit      := 0,    // 首扫态：输出直接采样输入，历史状态清零并置重算标记 / First scan: output tracks input, history cleared, recalc flagged
    eCoeffCalc := 10,   // 系数重算态：双线性变换重算五系数，检查钳位 / Coefficient recalc: bilinear recompute of five coefficients with clamping
    eRun       := 20,   // 运行态：双二阶递推滤波，系数保持不变 / Running: biquad recursion with unchanged coefficients
    eTrack     := 30,   // 跟踪态：输出立即跟随跟踪值，全部历史同步清零 / Tracking: output follows track value, all history synchronized to zero
    eFault     := 99    // 故障兜底态：非法状态进入，输出安全值并置故障码 / Fault fallback: entered from illegal states, safe output plus error code
);
END_TYPE

(*==============================================================================
 * 功能块: FB_DL_SecondOrderFilter
 * 调用约定: 每个采样周期无条件调用一次；fCutoffFreq 运行中可调，变更拍
 *           自动重算系数；tSampleTime 由调用方显式给定，不得依赖隐式扫描周期。
 * 滞后披露: 截止频率处幅值衰减约 -3dB、相位滞后约 90 度；等效群延迟随
 *           fCutoffFreq/fDt 比值变化，选型时需保证截止频率远低于奈奎斯特频率。
 * 递推披露: 采用双二阶直接型递推（输入历史 + 输出状态），与规格书公式
 *           fOut := fB0*fIn + fB1*fIn1 + fB2*fIn2 - fA1*fW1 - fA2*fW2 一致，
 *           fW1/fW2 承载上两拍输出状态，数学上与 II 型实现传递函数等价。
 *============================================================================*)
FUNCTION_BLOCK FB_DL_SecondOrderFilter
VAR_INPUT
    bEnable     : BOOL := FALSE;      // 使能，FALSE 时输出直通原始输入 / Enable, FALSE passes raw input straight through
    fIn         : REAL := 0.0;        // 原始采样输入 [EU] / Raw sampling input [EU]
    fCutoffFreq : REAL := 5.0;        // 截止频率 [Hz]，大于 0 且低于 0.45 倍采样频率 / Cutoff frequency [Hz], positive and below 0.45 times sampling rate
    bTrack      : BOOL := FALSE;      // 跟踪使能，TRUE 时输出立即跟随跟踪值 / Track enable, TRUE makes output follow track value instantly
    fTrackValue : REAL := 0.0;        // 跟踪目标值 [EU]，无扰投切用 / Track target value [EU], for bumpless transfer
    tSampleTime : TIME := T#100MS;    // 采样周期，小于 10ms 钳位 / Sampling period, clamped to 10ms minimum
END_VAR
VAR_OUTPUT
    fOut        : REAL;               // 滤波输出 [EU] / Filtered output [EU]
    bCoeffValid : BOOL;               // 系数就绪标志，重算完成置 TRUE / Coefficient ready flag, TRUE after recalculation
    bValid      : BOOL;               // 输出有效标志 / Output valid flag
    bError      : BOOL;               // 故障标志，与 uErrorId 联动 / Fault flag, coupled with uErrorId
    uErrorId    : UDINT;              // 故障码，0 = 无故障 / Error code, 0 = no error
END_VAR
VAR
    fB0         : REAL := 1.0;        // 递推系数 b0 [1]，初始为直通 / Recursion coefficient b0, initialized as pass-through
    fB1         : REAL := 0.0;        // 递推系数 b1 [1] / Recursion coefficient b1
    fB2         : REAL := 0.0;        // 递推系数 b2 [1] / Recursion coefficient b2
    fA1         : REAL := 0.0;        // 递推系数 a1 [1] / Recursion coefficient a1
    fA2         : REAL := 0.0;        // 递推系数 a2 [1] / Recursion coefficient a2
    fIn1        : REAL := 0.0;        // 上拍输入历史 [EU] / Previous input history [EU]
    fIn2        : REAL := 0.0;        // 上上拍输入历史 [EU] / Input history of two cycles ago [EU]
    fW1         : REAL := 0.0;        // 输出状态变量（上拍输出）[EU] / Output state variable (previous output) [EU]
    fW2         : REAL := 0.0;        // 输出状态变量（上上拍输出）[EU] / Output state variable (output two cycles ago) [EU]
    fDt         : REAL;               // 采样周期秒值 [s] / Sampling period in seconds [s]
    fFs         : REAL;               // 采样频率 [Hz] / Sampling frequency [Hz]
    fCutoffEff  : REAL;               // 钳位后的生效截止频率 [Hz] / Effective clamped cutoff frequency [Hz]
    fCutoffPrev : REAL := -1.0;       // 上次重算所用截止频率，用于变更检测 [Hz] / Cutoff used at last recalc, for change detection [Hz]
    fDtPrev     : REAL := -1.0;       // 上次重算所用周期，用于变更检测 [s] / Period used at last recalc, for change detection [s]
    fWc         : REAL;               // 归一化数字角频率 [rad] / Normalized digital angular frequency [rad]
    fK          : REAL;               // 预畸变中间量 tan(fWc/2) [1] / Prewarping intermediate tan(fWc/2) [1]
    fNorm       : REAL;               // 归一化分母 [1] / Normalization denominator [1]
    bCoeffDirty : BOOL := TRUE;       // 参数变更标记，TRUE 触发重算 / Parameter change flag, TRUE triggers recalculation
    eState      : E_DL_SofState;      // 状态机当前状态 / Current state of the state machine
END_VAR
VAR CONSTANT
    DL_SOF_SQRT2    : REAL := 1.4142136;  // 二阶巴特沃斯阻尼项系数根号二 [1] / Butterworth damping term sqrt(2) [1]
    DL_SOF_PI       : REAL := 3.1415927;  // 圆周率 [rad] / Pi constant [rad]
    DL_SOF_FC_MIN   : REAL := 1.0;        // 截止频率防御下限 [Hz] / Defensive cutoff frequency lower bound [Hz]
    DL_SOF_NYQ_KEEP : REAL := 0.45;       // 奈奎斯特保持系数（钳位到 0.45 倍采样频率）[1] / Nyquist keep ratio, clamp at 0.45 times sampling rate [1]
    DL_SOF_TAN_MAX  : REAL := 1.55;       // TAN 自变量上限 [rad]，防逼近奇异点 / TAN argument upper bound [rad], away from singularity
    DL_SOF_DT_MIN   : REAL := 0.01;       // 采样周期防御下限 [s] / Defensive sampling period lower bound [s]
    DL_SOF_INF_MAX  : REAL := 1.0E30;     // 有限值判定幅值上限 [EU] / Magnitude bound for finite-value check [EU]
END_VAR

(*------------------------------------------------------------------------------
 * 段 1｜采样周期钳位与派生量：dt 下限保护，采样频率反算
 *      Sampling period clamping and derived quantities
 *-----------------------------------------------------------------------------*)
uErrorId := 16#0002_0000;

IF tSampleTime < T#10MS THEN
    fDt      := DL_SOF_DT_MIN;                       // 周期过小钳位到 10ms / Too small period clamped to 10ms
    uErrorId := 16#0002_0002;                        // 采样周期非法已钳位 / Invalid sampling period clamped
ELSE
    fDt := TIME_TO_REAL(tSampleTime) / 1000.0;       // TIME 换算秒值 / Convert TIME to seconds
END_IF

fFs := 1.0 / fDt;                                    // 采样频率反算，fDt 已有下限保证 / Sampling frequency, guaranteed by dt floor

(*------------------------------------------------------------------------------
 * 段 2｜参数变更检测（浮点容差比较，禁止判等）：变更则置重算标记
 *      Parameter change detection with float tolerance, never equality
 *-----------------------------------------------------------------------------*)
IF (ABS(fCutoffFreq - fCutoffPrev) > 1.0E-6) OR (ABS(fDt - fDtPrev) > 1.0E-6) THEN
    bCoeffDirty := TRUE;                             // 截止频率或周期变更，触发重算 / Cutoff or period changed, trigger recalculation
END_IF

(*------------------------------------------------------------------------------
 * 段 3｜非有限值防御：拒绝本拍更新、保持上一拍输出（公共故障码）
 *      Non-finite defense: reject this cycle, hold previous output
 *-----------------------------------------------------------------------------*)
IF (fIn <> fIn) OR (ABS(fIn) > DL_SOF_INF_MAX) THEN
    uErrorId := 16#0002_0004;                        // 输入非有限值已拒绝 / Non-finite input rejected
    bValid   := FALSE;
    bError   := TRUE;
    RETURN;
END_IF

(*------------------------------------------------------------------------------
 * 段 4｜主状态机（红线 R6）：ENUM + CASE + ELSE 兜底
 *      Main state machine with mandatory ELSE fallback
 *-----------------------------------------------------------------------------*)
IF bTrack THEN
    eState := eTrack;                                // 跟踪请求优先级最高 / Track request has highest priority
ELSIF eState = eInit THEN
    eState := eInit;                                 // 首扫先采样直通，防首拍输出跳零 / First scan samples directly, no zero jump
ELSIF bCoeffDirty THEN
    eState := eCoeffCalc;                            // 参数变更进入重算态 / Parameter change enters recalc state
ELSIF eState = eFault THEN
    IF NOT bEnable THEN
        eState := eInit;                             // 使能跌落提供故障恢复路径 / Disabled input provides fault recovery path
    ELSE
        eState := eFault;                            // 故障态保持直至调用方处置 / Fault state holds until caller intervenes
    END_IF
ELSE
    eState := eRun;                                  // 常规运行态派生 / Normal running state derived
END_IF

CASE eState OF

    eInit:
        (* 首扫直接采样：历史清零并置重算标记，下一拍进入系数重算 *)
        (* First scan samples directly: history cleared and recalc flagged *)
        fOut        := fIn;
        fIn1        := fIn;
        fIn2        := fIn;
        fW1         := 0.0;
        fW2         := 0.0;
        bCoeffValid := FALSE;
        bValid      := FALSE;                        // 首扫未完成，输出尚不可信 / First scan unfinished, output not trustworthy yet
        bCoeffDirty := TRUE;
        eState      := eCoeffCalc;                   // 下一拍重算系数，避免系数未就绪递推 / Recalculate coefficients next cycle

    eCoeffCalc:
        (* 系数重算态：截止频率钳位 + 双线性变换预畸变 + 五系数归一化 *)
        (* Coefficient recalc: cutoff clamping, bilinear prewarping, normalization *)
        IF fCutoffFreq <= 0.0 THEN
            fCutoffEff := DL_SOF_FC_MIN;                 // 非法截止频率钳位到 1Hz / Illegal cutoff clamped to 1Hz
            uErrorId   := 16#0002_1101;                  // 截止频率非法已钳位 / Invalid cutoff frequency clamped
        ELSIF fCutoffFreq >= (fFs * 0.5) THEN
            fCutoffEff := fFs * DL_SOF_NYQ_KEEP;         // 越奈奎斯特钳位到 0.45 倍采样频率 / Over-Nyquist clamped to 0.45 times rate
            uErrorId   := 16#0002_1101;                  // 截止频率超奈奎斯特已钳位 / Cutoff over Nyquist clamped
        ELSE
            fCutoffEff := fCutoffFreq;                   // 合法参数原值生效 / Valid parameter applied as-is
        END_IF

        (* 归一化数字角频率与预畸变：TAN 自变量钳位防逼近奇异点 *)
        (* Normalized angular frequency with TAN argument clamped away from singularity *)
        fWc   := 2.0 * DL_SOF_PI * fCutoffEff * fDt;     // 数字角频率 [rad] / Digital angular frequency [rad]
        fK    := TAN(MIN(fWc / 2.0, DL_SOF_TAN_MAX));    // 预畸变中间量 / Prewarping intermediate value
        fNorm := 1.0 + DL_SOF_SQRT2 * fK + fK * fK;      // 归一化分母，恒大于零 / Normalization denominator, always positive

        IF ABS(fNorm) < 1.0E-9 THEN
            (* 分母退化防御（数学上不可达，防御性双检）：退化为直通系数 *)
            (* Degenerate denominator guard (mathematically unreachable): pass-through fallback *)
            fB0 := 1.0;
            fB1 := 0.0;
            fB2 := 0.0;
            fA1 := 0.0;
            fA2 := 0.0;
        ELSE
            (* 巴特沃斯五系数：直流增益经归一化恒为 1.000000 *)
            (* Butterworth coefficients: DC gain normalized to exactly 1.000000 *)
            fB0 := fK * fK / fNorm;
            fB1 := 2.0 * fB0;
            fB2 := fB0;
            fA1 := 2.0 * (fK * fK - 1.0) / fNorm;
            fA2 := (1.0 - DL_SOF_SQRT2 * fK + fK * fK) / fNorm;
        END_IF

        fCutoffPrev  := fCutoffEff;                  // 记录重算口径，供变更检测比对 / Record recalc baseline for change detection
        fDtPrev      := fDt;
        bCoeffValid  := TRUE;
        bCoeffDirty  := FALSE;
        eState       := eRun;

    eTrack:
        (* 无扰跟踪：输出立即跟随跟踪值，全部递推历史同步清零，回自动无跳变 *)
        (* Bumpless tracking: output follows track value, all recursion history cleared *)
        fOut        := fTrackValue;
        fIn1        := fTrackValue;
        fIn2        := fTrackValue;
        fW1         := 0.0;
        fW2         := 0.0;
        bCoeffDirty := TRUE;                         // 回运行态前强制重算一次系数 / Force one recalculation before running
        bValid      := TRUE;
        eState      := eRun;

    eRun:
        IF NOT bEnable THEN
            (* 使能失效语义：直通原始输入，历史同步防止恢复使能时残留跳变 *)
            (* Disabled semantics: pass raw input, history synchronized to avoid resume jumps *)
            fOut   := fIn;
            fIn1   := fIn;
            fIn2   := fIn;
            fW1    := 0.0;
            fW2    := 0.0;
            bValid := FALSE;
        ELSE
            (* 双二阶递推：按规格书公式执行，fW1/fW2 为上两拍输出状态 *)
            (* Biquad recursion per spec formula, fW1/fW2 carry previous two outputs *)
            fOut := fB0 * fIn + fB1 * fIn1 + fB2 * fIn2 - fA1 * fW1 - fA2 * fW2;
            fIn2 := fIn1;                            // 输入历史右移一位 / Shift input history by one
            fIn1 := fIn;
            fW2  := fW1;                             // 输出状态右移一位 / Shift output state by one
            fW1  := fOut;
            bValid := TRUE;
        END_IF

    eFault:
        (* 故障兜底：输出保持安全值 0，等待调用方修正后经使能跌落恢复 *)
        (* Fault fallback: output holds safe value 0, recovers via disabled input *)
        fOut        := 0.0;
        bCoeffValid := FALSE;
        bValid      := FALSE;

    ELSE
        (* 非法状态拦截：任何未定义枚举值一律进故障态并置公共兜底码 *)
        (* Illegal state interception: undefined enum values go to fault with code *)
        eState   := eFault;
        fOut     := 0.0;
        bValid   := FALSE;
        uErrorId := 16#0002_0005;

END_CASE;

(* 故障标志统一出口：与故障码严格联动，0 即无故障 *)
(* Unified fault flag outlet: strictly coupled with error code, zero means healthy *)
bError := (uErrorId <> 16#0002_0000);
END_FUNCTION_BLOCK
